(* IEC 61131-3 sources: iecf/harness/cases (part 4) *)

(* ---- bitarith.st ---- *)
(* Arithmetic on bit strings (the bit-string-arithmetic extension): a
   bit string counts as the unsigned integer of its width. Worked by
   hand, d 16#FFFF_FFF0, w 300, b 200, b2 100, i -5, x 513.7:
   %QD0  d + 16#20: DWORD, 16#1_0000_0010 wraps to 16#10, flagged.
   %QW4  w * 2 + b: WORD, 800 (16#0320); b widens to WORD.
   %QB6  b + b2: BYTE, 300 wraps to 44 (16#2C), flagged.
   %QW8  i + b: INT, -5 + 200 = 195; b counts as USINT, which INT holds.
   %QD12 BYTE_TO_REAL(b) + WORD_TO_REAL(w) / 3.0: 200.0 + 100.0 = 300.0
         (16#43960000), by value.
   %QB16 REAL_TO_BYTE(x / 10.0): 51.37 rounds to 51 (16#33).
   %QW18 w MOD 7 + b / 3: WORD 6 and BYTE 66 (division toward 0), as
         WORD 72 (16#48), into a UINT.
   %QB20 b - b2 * 2: 200 - 200 = 0.
   %QW22 a[b]: the array indexed by a BYTE, a[200] = 7.
   %QD24 DWORD_TO_REAL(16#3F800000) > 0.5: Ed.3's binary transfer is
         kept, 1.0 > 0.5, TRUE, 1.
   reference-skip: arithmetic on bit strings is CODESYS's, not IEC 61131-3. *)
PROGRAM main
  VAR
    d : DWORD := 16#FFFF_FFF0; w : WORD := 300; b : BYTE := 200; b2 : BYTE := 100;
    i : INT := -5; x : REAL := 513.7;
    a : ARRAY[0..255] OF INT;
  END_VAR
  VAR
    q0 AT %QD0 : DWORD; q1 AT %QW4 : WORD; q2 AT %QB6 : BYTE; q3 AT %QW8 : INT;
    q4 AT %QD12 : REAL; q5 AT %QB16 : BYTE; q6 AT %QW18 : UINT; q7 AT %QB20 : BYTE;
    q8 AT %QW22 : INT; q9 AT %QD24 : DWORD;
  END_VAR
  a[b] := 7;
  q0 := d + 16#20;
  q1 := w * 2 + b;
  q2 := b + b2;
  q3 := i + b;
  q4 := BYTE_TO_REAL(b) + WORD_TO_REAL(w) / 3.0;
  q5 := REAL_TO_BYTE(x / 10.0);
  q6 := w MOD 7 + b / 3;
  q7 := b - b2 * 2;
  q8 := a[b];
  q9 := DWORD_TO_REAL(16#3F800000) > 0.5;
END_PROGRAM

CONFIGURATION cf
  RESOURCE r ON x
    TASK tk(INTERVAL := T#10ms, PRIORITY := 1);
    PROGRAM p WITH tk : main;
  END_RESOURCE
END_CONFIGURATION

(* ---- bits.st ---- *)
(* Bit strings and BOOL: AND OR XOR NOT, the shifts and rotations, and
   BOOL expressions with short and full evaluation alike. *)
PROGRAM main
VAR
  x AT %IW0 : WORD;
  n AT %IB2 : BYTE;
  b0 AT %IX3.0 : BOOL;
  b1 AT %IX3.1 : BOOL;
  r_and AT %MW0 : WORD;
  r_or AT %MW2 : WORD;
  r_xor AT %MW4 : WORD;
  r_not AT %MW6 : WORD;
  r_shl AT %MW8 : WORD;
  r_shr AT %MW10 : WORD;
  r_rol AT %MW12 : WORD;
  r_ror AT %MW14 : WORD;
  r_dw AT %MD16 : DWORD;
  r_lw AT %ML20 : LWORD;
  r_by AT %MB28 : BYTE;
  q0 AT %QX0.0 : BOOL;
  q1 AT %QX0.1 : BOOL;
  q2 AT %QX0.2 : BOOL;
  q3 AT %QX0.3 : BOOL;
  q4 AT %QX0.4 : BOOL;
END_VAR
r_and := x AND 16#0FF0;
r_or := x OR 16#8001;
r_xor := x XOR 16#FFFF;
r_not := NOT x;
r_shl := SHL(x, BYTE_TO_INT(n));
r_shr := SHR(x, BYTE_TO_INT(n));
r_rol := ROL(x, BYTE_TO_INT(n));
r_ror := ROR(x, BYTE_TO_INT(n));
r_dw := ROL(WORD_TO_DWORD(x), 20);
r_lw := SHL(WORD_TO_LWORD(x), 48) OR 16#FF;
r_by := NOT n XOR 16#0F;
q0 := b0 AND b1;
q1 := b0 OR b1;
q2 := b0 XOR b1;
q3 := NOT b0 & b1;
q4 := (b0 OR NOT b1) AND x <> 0;
END_PROGRAM

CONFIGURATION plant
  RESOURCE r ON PLC
    TASK fast(INTERVAL := T#10ms, PRIORITY := 0);
    PROGRAM p WITH fast : main;
  END_RESOURCE
END_CONFIGURATION

(* ---- caseany.st ---- *)
(* CASE on a selector of any elementary type (Ed.3 7.3.3.3.3: "a
   variable of elementary data type", its labels "literals, enumerated
   values, or subranges" it can be compared with): BOOL, the bit
   strings, CHAR and WCHAR, STRING and WSTRING, REAL, TIME, DATE and
   TOD; labels that are literals, constants and subranges; a selector
   that is a FUNCTION with effects, called once. q[i] is the arm taken,
   9 for ELSE. Worked by hand:

   tick 0, n 1: b TRUE 1; w 16#2 1; bb 1 1; lw 1 ELSE 9; 'a' 1; "a" 1;
   'ab' 1; "ab" 1; 1.0 1; T#1s 1; the date 1; noon 1. calls 1 (Q12).
   tick 1, n 2: b FALSE 2; w 16#4, in 4..8, 2; bb 2 ELSE 9; lw 2 1; 'c'
   in 'b'..'d' 2; "z" in "y".."z" 2; 'cd', the constant, 2; "zz" 2; 2.5
   in 2.0..3.0 2; T#3s in the constant 2s..5s 2; June in February to
   December 2; 13:30 2. calls 2.
   tick 2, n 3: b TRUE 1; w 16#8 2; bb 3 1; lw 3 9; 'x' 9; "q" 9; 'zz'
   in 'x'..'zzzz' 3; "q" 9; -1.0 9; T#9s 9; 2021 9; 01:00 9. calls 3.
   reference-skip: CASE on anything but an integer or an enumeration:
   refused. *)
FUNCTION bump : STRING[4]
  VAR_INPUT s : STRING[4]; END_VAR
  VAR_EXTERNAL calls : USINT; END_VAR
  calls := calls + 1;
  bump := s;
END_FUNCTION
PROGRAM main
  VAR CONSTANT kc : CHAR := 'b'; ks : STRING[4] := 'cd'; kt : TIME := T#2s; END_VAR
  VAR_EXTERNAL calls : USINT; END_VAR
  VAR b : BOOL; w : WORD; bb : BYTE; c : CHAR; s : STRING[4]; r : REAL; t : TIME; d : DATE; wc : WCHAR; lw : LWORD; ws : WSTRING[4]; tod1 : TOD; n : USINT; END_VAR
  VAR q AT %QB0 : ARRAY [0..11] OF USINT; qc AT %QB12 : USINT; END_VAR
  n := n + 1;
  b := (n MOD 2) = 1;
  w := SHL(WORD#1, n);
  bb := USINT_TO_BYTE(n);
  lw := USINT_TO_LWORD(n);
  CASE n OF 1: c := 'a'; s := 'ab'; wc := "a"; ws := "ab"; r := 1.0; t := T#1s; d := D#2020-01-01; tod1 := TOD#12:00:00;
            2: c := 'c'; s := 'cd'; wc := "z"; ws := "zz"; r := 2.5; t := T#3s; d := D#2020-06-15; tod1 := TOD#13:30:00;
  ELSE c := 'x'; s := 'zz'; wc := "q"; ws := "q"; r := -1.0; t := T#9s; d := D#2021-01-01; tod1 := TOD#01:00:00;
  END_CASE;
  CASE b OF TRUE: q[0] := 1; FALSE: q[0] := 2; END_CASE;
  CASE w OF 16#0002: q[1] := 1; 16#0004..16#0008: q[1] := 2; ELSE q[1] := 3; END_CASE;
  CASE bb OF 16#01, 16#03: q[2] := 1; ELSE q[2] := 9; END_CASE;
  CASE lw OF 16#2: q[3] := 1; ELSE q[3] := 9; END_CASE;
  CASE c OF 'a': q[4] := 1; kc..'d': q[4] := 2; ELSE q[4] := 9; END_CASE;
  CASE wc OF "a": q[5] := 1; "y".."z": q[5] := 2; ELSE q[5] := 9; END_CASE;
  CASE bump(s) OF 'ab': q[6] := 1; ks: q[6] := 2; 'x'..'zzzz': q[6] := 3; ELSE q[6] := 9; END_CASE;
  CASE ws OF "ab": q[7] := 1; "zz": q[7] := 2; ELSE q[7] := 9; END_CASE;
  CASE r OF 1.0: q[8] := 1; 2.0..3.0: q[8] := 2; ELSE q[8] := 9; END_CASE;
  CASE t OF T#1s: q[9] := 1; kt..T#5s: q[9] := 2; ELSE q[9] := 9; END_CASE;
  CASE d OF D#2020-01-01: q[10] := 1; D#2020-02-01..D#2020-12-31: q[10] := 2; ELSE q[10] := 9; END_CASE;
  CASE tod1 OF TOD#12:00:00: q[11] := 1; TOD#13:00:00..TOD#14:00:00: q[11] := 2; ELSE q[11] := 9; END_CASE;
  qc := calls;
END_PROGRAM
CONFIGURATION c VAR_GLOBAL calls : USINT; END_VAR RESOURCE r ON PLC TASK t(INTERVAL := T#10ms, PRIORITY := 1); PROGRAM p WITH t : main; END_RESOURCE END_CONFIGURATION

(* ---- caselimits.st ---- *)
(* CASE subrange labels with a bound at the selector type's own limit:
   `0..5` on a USINT, `-128..-1` and `1..127` on a SINT, `0..255` on a
   USINT, all of it. Such a bound tests nothing, and its comparison is
   one C calls always true (-Wtype-limits): the generated C must still
   be strict-clean. Worked by hand, n and b counting 0, 1, 2 from tick 0,
   s -128, then -1, then 126:

   tick 0: n 0 in 0..5: Q0 01; s -128: Q1 01; b 0: Q2 01.
   tick 1: n 1: 01; s -1: 01; b 1: 01.
   tick 2: n 2: 01; s 126: Q1 03; 01. *)
PROGRAM main
  VAR n : USINT; s : SINT := -128; b : USINT; k : INT; END_VAR
  VAR q0 AT %QB0 : USINT; q1 AT %QB1 : USINT; q2 AT %QB2 : USINT; END_VAR
  CASE n OF 0..5: q0 := 1; ELSE q0 := 2; END_CASE;
  CASE s OF -128..-1: q1 := 1; 0: q1 := 2; 1..127: q1 := 3; END_CASE;
  CASE b OF 0..255: q2 := 1; END_CASE;
  n := n + 1;
  b := b + 1;
  k := k + 1;
  IF k = 1 THEN s := -1; ELSE s := 126; END_IF;
END_PROGRAM
CONFIGURATION c RESOURCE r ON PLC TASK t(INTERVAL := T#10ms, PRIORITY := 1); PROGRAM p WITH t : main; END_RESOURCE END_CONFIGURATION

(* ---- casenamed.st ---- *)
(* A named value as a CASE label (Ed.3 6.4.4.3, 7.3.3.3.3): a constant,
   its number compared with the selector's. Found in TcOpen, where it
   was E0032. Worked by hand:
   %QW0: d is eDist#Y (20): the label eDist#Y, 2.
   %QW2: n is eNum#Q (5): the label eNum#Q, 4.
   %QW4: d's number through its base type, 20.
   reference-skip: matiec has no named values with values given. *)
TYPE eDist : (X := 10, Y := 20, Z := 30); END_TYPE
TYPE eNum : INT (P := 1, Q := 5); END_TYPE

PROGRAM main
  VAR d : eDist := eDist#Y; n : eNum := eNum#Q; END_VAR
  VAR q0 AT %QW0 : INT; q1 AT %QW2 : INT; q2 AT %QW4 : INT; END_VAR
  CASE d OF
    eDist#X: q0 := 1;
    eDist#Y: q0 := 2;
  ELSE
    q0 := 3;
  END_CASE;
  CASE n OF
    eNum#P: q1 := 3;
    eNum#Q: q1 := 4;
  END_CASE;
  q2 := TO_INT(d);
END_PROGRAM

CONFIGURATION cf
  RESOURCE r ON x
    TASK tk(INTERVAL := T#10ms, PRIORITY := 1);
    PROGRAM p WITH tk : main;
  END_RESOURCE
END_CONFIGURATION

(* ---- codesysanyto.st ---- *)
(* CODESYS's and TwinCAT's ANY_TO_<type> (any-to): Ed.3's overloaded
   TO_<type>, as TcOpen's TcoRealToBytes and StringBuilder call it.
   Worked by hand, d + 1 and b + 1 each tick, d from 41, b from 7:
   %QW0 ANY_TO_INT(r * 2.0), r = ANY_TO_REAL(d): tick 0 d 42: 84;
   %QW2 ANY_TO_INT(ANY_TO_STRING(b) + '0' joined): b 7: '70': 70;
   %QW4 ANY_TO_INT(ANY_TO_BOOL(b - 7)): b 7: FALSE: 0.
   tick 1: d 43: 86; b 8: 80; 1.
   reference-skip: not IEC 61131-3. *)
PROGRAM main
  VAR d : DINT := 41; r : REAL; b : BYTE := 7; END_VAR
  VAR q0 AT %QW0 : INT; END_VAR
  VAR q1 AT %QW2 : INT; END_VAR
  VAR q2 AT %QW4 : INT; END_VAR
  d := d + 1;
  r := ANY_TO_REAL(d);
  q0 := ANY_TO_INT(r * 2.0);
  q1 := ANY_TO_INT(CONCAT(ANY_TO_STRING(b), '0'));
  q2 := ANY_TO_INT(ANY_TO_BOOL(b - 7));
  b := b + 1;
END_PROGRAM

CONFIGURATION cf
  RESOURCE r ON x
    TASK tk(INTERVAL := T#10ms, PRIORITY := 1);
    PROGRAM p WITH tk : main;
  END_RESOURCE
END_CONFIGURATION

(* ---- codesyschain.st ---- *)
(* Found in OSCAT BUILDING (BOILER): chained assignment, read right to
   left, each inner target read back (chained-assignment). Worked by hand:
   %QD0: r := x := 7 / 2: x is INT, 7 / 2 is 3, r gets 3.0, 16#40400000.
   %QW4: x, 3.
   %QW6, %QW8: q := arr[i] := y := 9, i 2: arr[2] 9, q 9.
   %QW10: inside IF, a := b := c := 5 then a + b + c: 15.
   reference-skip: not IEC 61131-3. *)
PROGRAM main
  VAR
    x : INT; y : SINT; i : INT := 2; arr : ARRAY[0..3] OF INT;
    a : INT; b : INT; c : INT;
  END_VAR
  VAR
    r AT %QD0 : REAL; qx AT %QW4 : INT; q AT %QW6 : INT; q2 AT %QW8 : INT;
    q3 AT %QW10 : INT;
  END_VAR
  r := x := 7 / 2;
  qx := x;
  q := arr[i] := y := 9;
  q2 := arr[2];
  IF i = 2 THEN
    a := b := c := 5;
  END_IF;
  q3 := a + b + c;
END_PROGRAM

CONFIGURATION cf
  RESOURCE r ON x
    TASK tk(INTERVAL := T#10ms, PRIORITY := 1);
    PROGRAM p WITH tk : main;
  END_RESOURCE
END_CONFIGURATION

(* ---- codesysdates.st ---- *)
(* Found in OSCAT NETWORK and BUILDING, each an extension. Worked by hand:
   %QB0 bit 0: UDINT 70000 > DWORD 16#10000 (65536): a bit string compared
   with an integer, as its unsigned integer (bit-string-arithmetic): TRUE.
   %QB0 bit 1: BYTE 200 < INT 100: FALSE.
   %QW2: TOD_TO_TIME(TOD#01:00:00) is T#1h, as DINT ms / 1000, 3600.
   %QD4: TIME_TO_TOD(T#1d2h3m4s5ms) drops the day: TOD#02:03:04.005,
   7384005 ms (date-number-conversions).
   %QD8: D#2026-11-19 + T#1d - T#2d is D#2026-11-18; DATE_TO_UDINT /
   86400 counts its days since 1970-01-01: 20775
   (date-time-arithmetic).
   %QB12: d2 := d + half, half T#12h a variable: no whole day, flagged
   and left undone, d2 stays D#1970-01-01: DATE_TO_UDINT(d2) = 0.
   reference-skip: none of these is IEC 61131-3. *)
PROGRAM main
  VAR
    u : UDINT := 70000; w : DWORD := 16#10000; b : BYTE := 200; i : INT := 100;
    d : DATE := D#2026-11-19; d2 : DATE; half : TIME := T#12h;
  END_VAR
  VAR
    x0 AT %QX0.0 : BOOL; x1 AT %QX0.1 : BOOL; q1 AT %QW2 : INT; q2 AT %QD4 : UDINT;
    q3 AT %QD8 : UDINT; q4 AT %QB12 : BYTE;
  END_VAR
  x0 := u > w;
  x1 := b < i;
  q1 := DINT_TO_INT(TIME_TO_DINT(TOD_TO_TIME(TOD#01:00:00)) / 1000);
  q2 := TOD_TO_UDINT(TIME_TO_TOD(T#1d2h3m4s5ms));
  q3 := DATE_TO_UDINT(d + T#1d - T#2d) / 86400;
  d2 := d + half;
  q4 := UDINT_TO_BYTE(DATE_TO_UDINT(d2));
END_PROGRAM

CONFIGURATION cf
  RESOURCE r ON x
    TASK tk(INTERVAL := T#10ms, PRIORITY := 1);
    PROGRAM p WITH tk : main;
  END_RESOURCE
END_CONFIGURATION

(* ---- codesysdtliterals.st ---- *)
(* A DT literal's seconds left out, and a fraction of its second
   (dt-literals): the seconds 0, the fraction dropped, W0016 - as
   TcOpen's TcoMessenger writes DT#1970-01-01-00:00 and its
   fbManipulatorAutomat DT#2013-05-09-13:29:20.500. Worked by hand,
   each as its seconds since 1970 (date-number-conversions):
   DT#1970-01-01-00:01: 60, 16#3C (%QD0).
   DT#2013-05-09-13:29:20.500: 2013-05-09 is day 15834, 1368057600 s;
   13:29:20 is 48560 s; 1368106160, 16#518BA4B0 (%QD4).
   An initial value DT#1970-01-02-00:00:00.999: one day, 86400, 16#15180
   (%QD8).
   reference-skip: not IEC 61131-3. *)
PROGRAM main
  VAR
    a : DT; b : DT; c : DT := DT#1970-01-02-00:00:00.999;
  END_VAR
  VAR q0 AT %QD0 : UDINT; q1 AT %QD4 : UDINT; q2 AT %QD8 : UDINT; END_VAR
  a := DT#1970-01-01-00:01;
  b := DT#2013-05-09-13:29:20.500;
  q0 := DT_TO_UDINT(a);
  q1 := DT_TO_UDINT(b);
  q2 := DT_TO_UDINT(c);
END_PROGRAM

CONFIGURATION cf
  RESOURCE r ON x
    TASK tk(INTERVAL := T#10ms, PRIORITY := 1);
    PROGRAM p WITH tk : main;
  END_RESOURCE
END_CONFIGURATION

(* ---- codesysenum.st ---- *)
(* CODESYS's enumerations (the codesys-enums extension,
   docs/extensions.md): the base type after the values, `(...) DWORD :=
   black`, and a value named `COLOR.green`, as CODESYS and TwinCAT write
   them (their `qualified_only` makes every use so); the attributes
   before a TYPE are pragmas, which iecf reads past. Worked by hand:
   COLOR is DWORD, black its initial value: c is 16#88000000, its top
   byte 16#88 (%QB0); c := COLOR.green, 16#FF00FF00, top byte 16#FF
   (%QB1); c = COLOR.green TRUE (%QX4.0). Lib.Mode (stop, run, fault)
   starts as Lib.Mode.stop: m = Lib.Mode.stop, 1 at tick 0, then 0
   (%QB2); m := Lib.Mode.run; CASE m OF Lib.Mode.run: %QB3 := 7.
   reference-skip: CODESYS's writing is not IEC 61131-3. *)
{attribute 'qualified_only'}
{attribute 'strict'}
TYPE COLOR :
(
    white := 16#FFFFFF00,
    green := 16#FF00FF00,
    black := 16#88000000
) DWORD := black
;
END_TYPE

NAMESPACE Lib
  TYPE Mode : (stop, run, fault); END_TYPE
END_NAMESPACE

PROGRAM main
  VAR c : COLOR; m : Lib.Mode := Lib.Mode.stop; END_VAR
  VAR
    q0 AT %QB0 : BYTE;
    q1 AT %QB1 : BYTE;
    q2 AT %QB2 : SINT;
    q3 AT %QB3 : SINT;
    b0 AT %QX4.0 : BOOL;
  END_VAR
  c := COLOR#black;
  q0 := DWORD_TO_BYTE(SHR(c, 24));
  c := COLOR.green;
  q1 := DWORD_TO_BYTE(SHR(c, 24));
  b0 := c = COLOR.green;
  q2 := SEL(m = Lib.Mode.stop, SINT#0, SINT#1);
  m := Lib.Mode.run;
  CASE m OF
    Lib.Mode.stop: q3 := 1;
    Lib.Mode.run: q3 := 7;
  END_CASE;
END_PROGRAM

CONFIGURATION cf
  RESOURCE r ON x
    TASK t(INTERVAL := T#10ms, PRIORITY := 1);
    PROGRAM p WITH t : main;
  END_RESOURCE
END_CONFIGURATION

(* ---- codesysgvl.st ---- *)
(* Global variable lists (--gvl, --qualified-gvl), as CODESYS and TwinCAT
   name them: IO (codesysgvl.d/io.st) and CFG, qualified-only
   (codesysgvl.d/cfg.st). Worked by hand:
   cycle 0: %QW0 IO.a + CFG.k = 3 + 7 = 10; r[CFG.N] := IO.a, %QW2 3;
     IO.a 4, read bare: %QW4 4; CFG.t[4] := 4 + 1, %QW6 5.
   cycle 1: 4 + 7 = 11; 4; 5; 6.
   reference-skip: not IEC 61131-3. *)
PROGRAM main
  VAR r : ARRAY[1..CFG.N] OF INT; END_VAR
  VAR x AT %QW0 : INT; y AT %QW2 : INT; z AT %QW4 : INT; w AT %QW6 : INT; END_VAR
  x := IO.a + CFG.k;
  r[CFG.N] := IO.a;
  y := r[4];
  IO.a := IO.a + 1;
  z := a;
  CFG.t[CFG.N] := a + 1;
  w := CFG.t[4];
END_PROGRAM

CONFIGURATION cf
  RESOURCE r ON x
    TASK tk(INTERVAL := T#10ms, PRIORITY := 1);
    PROGRAM p WITH tk : main;
  END_RESOURCE
END_CONFIGURATION

(* ---- codesysjump.st ---- *)
(* Found in OSCAT NETWORK (IP_CONTROL2): JMP and labels in ST
   (jump-labels). Worked by hand:
   %QW0: i counted to 5 by a jump back: 5.
   %QW2: JMP out of the FOR at k = 3, k left as the body has it: 3.
   %QW4: n = 1 + 2 + 3: 6; the jumped-over q2 := 99 never runs.
   %QW6: arr[k] with k 2 holds; k 7 on the jump back is outside 0..3:
   INDEX fault on the line of arr[k] := 1 (32), the task stops: q3 1.
   reference-skip: not IEC 61131-3. *)
PROGRAM main
  VAR i : INT; k : INT; n : INT; arr : ARRAY[0..3] OF INT; END_VAR
  VAR q0 AT %QW0 : INT; q1 AT %QW2 : INT; q2 AT %QW4 : INT; q3 AT %QW6 : INT; END_VAR
  i := 0;
  n := 0;
again:
  i := i + 1;
  IF i < 5 THEN
    JMP again;
  END_IF;
  q0 := i;
  JMP skip;
  q2 := 99;
skip:
  FOR k := 1 TO 10 DO
    n := n + k;
    IF k = 3 THEN JMP out; END_IF;
  END_FOR;
out:
  q1 := k;
  q2 := n;
  k := 2;
back:
  arr[k] := 1;
  k := k + 5;
  q3 := q3 + 1;
  IF k < 20 THEN JMP back; END_IF;
END_PROGRAM

CONFIGURATION cf
  RESOURCE r ON x
    TASK tk(INTERVAL := T#10ms, PRIORITY := 1);
    PROGRAM p WITH tk : main;
  END_RESOURCE
END_CONFIGURATION

(* ---- codesyslibprograms.st ---- *)
(* A library's PROGRAMs in its namespace, as CODESYS and TwinCAT have
   them: the library A (codesyslibprograms.d/a.st) and B, qualified-only
   (b.st), each with a MAIN of its own, beside this project's MAIN. A's
   Counter is called and read by its short name, through A's USING,
   from here and from A's own block User, and its method called;
   A.MAIN and B.MAIN by the library's name (program-instances).
   Worked by hand:
   cycle 0: Counter() v 10, %QW0 10; A.MAIN() n 1, %QW2 1; B.MAIN()
     x 100, %QW4 100; u(), Counter() again, %QW6 20; A.Counter.Bump(5),
     %QW8 25.
   cycle 1: 35; 2; 200; 45; 50.
   reference-skip: not IEC 61131-3. *)
PROGRAM MAIN
  VAR u : User; END_VAR
  VAR q0 AT %QW0 : INT; q1 AT %QW2 : INT; q2 AT %QW4 : INT; q3 AT %QW6 : INT; q4 AT %QW8 : INT; END_VAR
  Counter();
  q0 := Counter.v;
  A.MAIN();
  q1 := A.MAIN.n;
  B.MAIN();
  q2 := B.MAIN.x;
  u();
  q3 := Counter.v;
  A.Counter.Bump(5);
  q4 := A.Counter.v;
END_PROGRAM

CONFIGURATION cf
  RESOURCE r ON x
    TASK tk(INTERVAL := T#10ms, PRIORITY := 1);
    PROGRAM p WITH tk : MAIN;
  END_RESOURCE
END_CONFIGURATION

(* ---- codesysliteralwidening.st ---- *)
(* An untyped integer literal the other operand's type does not hold
   (literal-widening): the operation is computed in the narrowest type
   of the operand's kind that holds it, as CODESYS and TwinCAT compute
   intermediate results at least 32 bits wide. TcOpen's TcoBytesToReal
   writes `256 * _b0 + _b1` of BYTEs and `w * 65536` of a WORD, its
   TcoRealToBytes `2147483648 + ...` of DINTs.
   Worked by hand:
   256 * 16#12 + 16#34, in WORD: 16#1234 (4660).
   16#0003 * 65536 + 16#1234, in DWORD: 16#00031234 (201268).
   2147483648 + 100, in LINT: 2147483748 (16#80000064).
   5 * -1 of a UINT, in DINT: -5.
   30000 < 70000 of an INT, compared in DINT: TRUE.
   reference-skip: not IEC 61131-3. *)
PROGRAM main
  VAR
    b0 : BYTE := 16#12;
    b1 : BYTE := 16#34;
    w : WORD;
    w1 : WORD := 16#0003;
    k : INT := 30000;
    x : DINT := 100;
    u : UINT := 5;
  END_VAR
  VAR q0 AT %QD0 : DWORD; q4 AT %QD4 : DWORD; q8 AT %QL8 : LINT; q16 AT %QD16 : DINT; q20 AT %QX20.0 : BOOL; END_VAR
  w := 256 * b0 + b1;
  q0 := w;
  q4 := (w1 * 65536) + w;
  q8 := 2147483648 + x;
  q16 := u * -1;
  q20 := k < 70000;
END_PROGRAM

CONFIGURATION cf
  RESOURCE r ON x
    TASK tk(INTERVAL := T#10ms, PRIORITY := 1);
    PROGRAM p WITH tk : main;
  END_RESOURCE
END_CONFIGURATION

(* ---- codesyspack.st ---- *)
(* The codesys pack (docs/extensions.md, "Packs"): one name for the
   extensions code written for CODESYS and TwinCAT uses, seven of them
   here. Worked by hand:
   gCount, a top-level global, used without VAR_EXTERNAL
   (implicit-externals) and bound to a REFERENCE TO (reference-to): r :=
   r + 1 makes it 6, then 7 (%QB3). t T#1500ms; ms := TIME_TO_DINT(t),
   1500 (time-number-conversions), worked out as it is set up
   (initial-expressions): ms / 100, 15 (%QB0). Len3 takes a VAR_IN_OUT
   CONSTANT STRING(10) (in-out-constant, string-parentheses), given 16
   characters, all of them read: n := Len3('abcdefghijklmnop') + ms,
   1516; n - 1500, 16 (%QB1). m : E_Mode := E_Mode.eRun, its base type
   after its values (codesys-enums): m = E_Mode.eRun, 1 (%QB2).
   BYTE_TO_BOOL(16#10) TRUE (bit-string-to-bool, %QX4.0).
   reference-skip: CODESYS's extensions are not IEC 61131-3. *)
VAR_GLOBAL gCount : INT := 5; END_VAR

TYPE E_Mode : (eIdle, eRun) DWORD; END_TYPE

FUNCTION Len3 : DINT
  VAR_IN_OUT CONSTANT s : STRING(10); END_VAR
  Len3 := INT_TO_DINT(LEN(s));
END_FUNCTION

PROGRAM main
  VAR
    t : TIME := T#1500ms;
    ms : DINT := TIME_TO_DINT(t);
    n : DINT := Len3('abcdefghijklmnop') + ms;
    m : E_Mode := E_Mode.eRun;
    r : REFERENCE TO INT;
    b : BOOL := BYTE_TO_BOOL(16#10);
  END_VAR
  VAR
    q0 AT %QB0 : SINT;
    q1 AT %QB1 : SINT;
    q2 AT %QB2 : SINT;
    q3 AT %QB3 : SINT;
    b0 AT %QX4.0 : BOOL;
  END_VAR
  r REF= gCount;
  r := r + 1;
  q0 := DINT_TO_SINT(ms / 100);
  q1 := DINT_TO_SINT(n - 1500);
  q2 := SEL(m = E_Mode.eRun, SINT#0, SINT#1);
  q3 := INT_TO_SINT(gCount);
  b0 := b;
END_PROGRAM

CONFIGURATION cf
  RESOURCE r ON x
    TASK tk(INTERVAL := T#10ms, PRIORITY := 1);
    PROGRAM p WITH tk : main;
  END_RESOURCE
END_CONFIGURATION

(* ---- codesyssemi.st ---- *)
(* Found in TcOpen (TwinCAT), 10639 ends without ';' against 829 with,
   and in OSCAT: END_IF and its kin with no ';' (optional-semicolons).
   Worked by hand:
   %QW0: n counts 1 + 2 + 3 + 4 by FOR, then +10 by IF: 20.
   %QW2: WHILE doubles w from 1 past 100: 128; REPEAT halves it to 64,
   then CASE adds 1 for 64: 65.
   reference-skip: not IEC 61131-3. *)
PROGRAM main
  VAR n : INT; i : INT; w : INT := 1; END_VAR
  VAR q0 AT %QW0 : INT; q1 AT %QW2 : INT; END_VAR
  n := 0;
  FOR i := 1 TO 4 DO
    n := n + i;
  END_FOR
  IF n = 10 THEN
    n := n + 10;
  END_IF
  WHILE w <= 100 DO
    w := w * 2;
  END_WHILE
  REPEAT
    w := w / 2;
  UNTIL w <= 100 END_REPEAT
  CASE w OF
    64: w := w + 1;
  END_CASE
  q0 := n;
  q1 := w;
END_PROGRAM

CONFIGURATION cf
  RESOURCE r ON x
    TASK tk(INTERVAL := T#10ms, PRIORITY := 1);
    PROGRAM p WITH tk : main;
  END_RESOURCE
END_CONFIGURATION

(* ---- codesysstraysemi.st ---- *)
(* A `;` that ends nothing (stray-semicolons), as TcOpen writes
   `END_TYPE;` after its EtherCAT structures and `p : T;;` in a VAR
   section; END_PROGRAM; too: dropped, the declarations read as
   without it.
   Worked by hand, each tick: s.a + 1 and s.b + 2 from 0; k counts.
   Tick 1: 1, 2, 1; tick 2: 2, 4, 2.
   reference-skip: not IEC 61131-3. *)
TYPE Pair :
STRUCT
  a : INT;
  b : INT;
END_STRUCT
END_TYPE;

PROGRAM main
  VAR
    s : Pair;;
    ;
    k : INT;
  END_VAR
  VAR q0 AT %QW0 : INT; q2 AT %QW2 : INT; q4 AT %QW4 : INT; END_VAR
  s.a := s.a + 1;
  s.b := s.b + 2;
  k := k + 1;
  q0 := s.a;
  q2 := s.b;
  q4 := k;
END_PROGRAM;

CONFIGURATION cf
  RESOURCE r ON x
    TASK tk(INTERVAL := T#10ms, PRIORITY := 1);
    PROGRAM p WITH tk : main;
  END_RESOURCE
END_CONFIGURATION

(* ---- codesysstructext.st ---- *)
(* A structure extending another (struct-extends), as TcOpen's I/O types
   do: TYPE X EXTENDS Base : STRUCT, the base's fields first, at any
   depth, their initial values with them. Worked by hand:
   %QW0: t.a := 1, then a + b + c + d: 1 + 2 + 3 + 4 = 10.
   %QW2: a Top given to a Middle's field by field: Middle.c, 3.
   reference-skip: not IEC 61131-3. *)
TYPE
  Base : STRUCT a : INT; b : INT := 2; END_STRUCT;
  Middle EXTENDS Base : STRUCT c : INT := 3; END_STRUCT;
  Top EXTENDS Middle : STRUCT d : INT := 4; END_STRUCT;
END_TYPE

PROGRAM main
  VAR t : Top; m : Middle; END_VAR
  VAR q AT %QW0 : INT; r AT %QW2 : INT; END_VAR
  t.a := 1;
  q := t.a + t.b + t.c + t.d;
  m.c := t.c;
  r := m.c;
END_PROGRAM

CONFIGURATION cf
  RESOURCE r ON x
    TASK tk(INTERVAL := T#10ms, PRIORITY := 1);
    PROGRAM p WITH tk : main;
  END_RESOURCE
END_CONFIGURATION

(* ---- codesyssyntax.st ---- *)
(* Three CODESYS ways of writing, each an extension (docs/extensions.md).
   Worked by hand:
   struct-semicolon: Pair ends END_STRUCT with no ';', the next type
   follows; Trio's END_STRUCT stands before END_TYPE.
   bare-array-init: a : ARRAY[1..5] OF SINT := 1, 2, 2(7), 3; is
   [1, 2, 7, 7, 3], sum 20 (%QB0); Pair's v := 8, 9 in a STRUCT, 8 + 9 =
   17 (%QB1); the type Row := 4, 5, 6, 4 + 5 + 6 = 15 (%QB2).
   real-without-point: r := 1E3 + 25E-1, 1002.5; REAL_TO_SINT(r / 100.0)
   is 10.025 rounded, 10 (%QB3); Trio's z := 2E1, 20.0, as SINT 20
   (%QB4).
   reference-skip: none of the three is IEC 61131-3. *)
TYPE
  Pair : STRUCT
    v : ARRAY[1..2] OF SINT := 8, 9;
  END_STRUCT
  Row : ARRAY[0..2] OF SINT := 4, 5, 6;
  Trio : STRUCT
    z : REAL := 2E1;
  END_STRUCT
END_TYPE

PROGRAM main
  VAR
    a : ARRAY[1..5] OF SINT := 1, 2, 2(7), 3;
    p : Pair;
    w : Row;
    t : Trio;
    r : REAL;
    i : INT;
    s : SINT;
  END_VAR
  VAR
    q0 AT %QB0 : SINT;
    q1 AT %QB1 : SINT;
    q2 AT %QB2 : SINT;
    q3 AT %QB3 : SINT;
    q4 AT %QB4 : SINT;
  END_VAR
  s := 0;
  FOR i := 1 TO 5 DO
    s := s + a[i];
  END_FOR;
  q0 := s;
  q1 := p.v[1] + p.v[2];
  q2 := w[0] + w[1] + w[2];
  r := 1E3 + 25E-1;
  q3 := REAL_TO_SINT(r / 100.0);
  q4 := REAL_TO_SINT(t.z);
END_PROGRAM

CONFIGURATION cf
  RESOURCE r ON x
    TASK tk(INTERVAL := T#10ms, PRIORITY := 1);
    PROGRAM p WITH tk : main;
  END_RESOURCE
END_CONFIGURATION

(* ---- codesysunion.st ---- *)
(* CODESYS's and TwinCAT's UNION (union), as a STRUCT OVERLAP whose every
   member is AT %B0: un set up through d alone, 1.0's bits (16#3F800000);
   r, declared first, is not defaulted over it. Worked by hand:
   %QD0: q := un.r before un.r is changed, 1.0's bytes, 00 00 80 3f.
   un.r := 2.0 changes the same bytes un.d reads.
   %QD4: w := un.d after that, 2.0's bits read as a DWORD, 00 00 00 40.
   reference-skip: not IEC 61131-3. *)
TYPE
  U : UNION
    r : REAL;
    d : DWORD;
  END_UNION;
END_TYPE

PROGRAM main
  VAR un : U := (d := 16#3F800000); END_VAR
  VAR q AT %QD0 : REAL; w AT %QD4 : DWORD; END_VAR
  q := un.r;
  un.r := 2.0;
  w := un.d;
END_PROGRAM

CONFIGURATION cf
  RESOURCE r ON x
    TASK tk(INTERVAL := T#10ms, PRIORITY := 1);
    PROGRAM p WITH tk : main;
  END_RESOURCE
END_CONFIGURATION

(* ---- connections.st ---- *)
(* Program connections (Ed.3 6.8.2): a program instance's inputs given a
   literal, a global or an address, its outputs written to a global or an
   address. Each input is set before the instance runs, each output
   taken after it. The reference compiler crashes on a literal input and writes C that
   does not compile for the rest (PROPOSAL.md §1b): the trace is iecf's
   alone, connections.iecf.trace, checked by hand.

   Instance a adds 1 a tick, b adds the global ten (10), c the input
   global k (at %IW0). a's total goes to the global sum, b's to the
   global out_b (at %MD4), c's to out_c (at %MD8); a's done, inverted,
   straight to the address %QX0.0, a bare BOOL. *)
PROGRAM counter
VAR_INPUT inc : INT; END_VAR
VAR_OUTPUT total : DINT; done : BOOL; END_VAR
total := total + inc;
done := total >= 3;
END_PROGRAM

PROGRAM report
VAR_EXTERNAL sum : DINT; END_VAR
VAR r_sum AT %MD0 : DINT; END_VAR
r_sum := sum;
END_PROGRAM

CONFIGURATION plant
  VAR_GLOBAL
    ten : INT := 10;
    sum : DINT;
  END_VAR
  VAR_GLOBAL
    k AT %IW0 : INT;
    out_b AT %MD4 : DINT;
    out_c AT %MD8 : DINT;
  END_VAR
  RESOURCE r ON PLC
    TASK fast(INTERVAL := T#10ms, PRIORITY := 0);
    PROGRAM a WITH fast : counter(inc := 1, total => sum, NOT done => %QX0.0);
    PROGRAM b WITH fast : counter(inc := ten, total => out_b);
    PROGRAM c WITH fast : counter(inc := k, total => out_c);
    PROGRAM rep WITH fast : report;
  END_RESOURCE
END_CONFIGURATION

(* ---- conrefs.st ---- *)
(* Program connections (Ed.3 6.8.2) of a reference, in and out, and of
   NULL; a CHAR output into a STRING global and a WCHAR one into a
   WSTRING global (Figure 11, implicit). The three programs run in
   order on one task. Worked by hand: setup points gr at gi (5). p1 gets
   gr, adds 1 to what it references and gives it back as ro, into gro;
   p2 gets NULL and does nothing, its ro NULL into gro2. Tick 0: gi 6
   (%QB0), gro^ 6 (%QB1), gro2 NULL (%QX2.0), gs 'k' (%QX2.1), gws "z"
   (%QX2.2). Tick 1: gi 7, gro^ 7.
   reference-skip: program connections, as connections; and REF_TO. *)
PROGRAM setup
  VAR_EXTERNAL gi : INT; gr : REF_TO INT; END_VAR
  gr := REF(gi);
END_PROGRAM

PROGRAM prod
  VAR_INPUT r : REF_TO INT; END_VAR
  VAR_OUTPUT ro : REF_TO INT; c : CHAR; wc : WCHAR; END_VAR
  IF r <> NULL THEN
    r^ := r^ + 1;
  END_IF;
  ro := r;
  c := 'k';
  wc := WCHAR#"z";
END_PROGRAM

PROGRAM show
  VAR_EXTERNAL gi : INT; gro, gro2 : REF_TO INT; gs : STRING[4]; gws : WSTRING[4]; END_VAR
  VAR
    q0 AT %QB0 : SINT;
    q1 AT %QB1 : SINT;
    b0 AT %QX2.0 : BOOL;
    b1 AT %QX2.1 : BOOL;
    b2 AT %QX2.2 : BOOL;
  END_VAR
  q0 := INT_TO_SINT(gi);
  IF gro <> NULL THEN
    q1 := INT_TO_SINT(gro^);
  END_IF;
  b0 := gro2 = NULL;
  b1 := gs = 'k';
  b2 := gws = "z";
END_PROGRAM

CONFIGURATION cf
  VAR_GLOBAL
    gi : INT := 5;
    gr, gro, gro2 : REF_TO INT;
    gs : STRING[4];
    gws : WSTRING[4];
  END_VAR
  RESOURCE r ON PLC
    TASK t(INTERVAL := T#10ms, PRIORITY := 1);
    PROGRAM s WITH t : setup;
    PROGRAM p1 WITH t : prod(r := gr, ro => gro, c => gs, wc => gws);
    PROGRAM p2 WITH t : prod(r := NULL, ro => gro2);
    PROGRAM v WITH t : show;
  END_RESOURCE
END_CONFIGURATION

(* ---- constinit2.st ---- *)
(* Initial values that are functions of constants (Table 34's string
   functions, the conversions of whole numbers to and from text, Tables
   30 and 36's date functions): worked out by the compiler. Each is
   compared with the same function of variables, computed as the program
   runs; ok counts those that agree, 19 of 19 (Q0 13). Worked by hand
   for three: LEN of s6, 'abZZef', is 6 (Q1); f1, FIND('abcabc', 'ca'),
   is 3 (Q2); i1, STRING_TO_INT('17'), is 17 (Q3 11).
   reference-skip: the reference compiler takes a literal there. *)
PROGRAM main
  VAR CONSTANT pre : STRING[4] := 'ab'; END_VAR
  VAR
    s1 : STRING[8] := CONCAT('ab', 'cd');
    s2 : STRING[8] := CONCAT(pre, '-x', 'y');
    l1 : INT := LEN('hello');
    s3 : STRING[8] := INT_TO_STRING(-42);
    s4 : STRING[8] := LEFT('abcdef', 3);
    s5 : STRING[8] := RIGHT('abcdef', 2);
    s6 : STRING[8] := REPLACE('abcdef', 'ZZ', 2, 3);
    s7 : STRING[8] := MID('abcdef', 2, 3);
    s9 : STRING[8] := INSERT('abcd', 'XY', 2);
    s10 : STRING[8] := DELETE('abcdef', 2, 3);
    ws : WSTRING[8] := CONCAT("ab", "cd");
    f1 : INT := FIND('abcabc', 'ca');
    i1 : INT := STRING_TO_INT('17');
    d1 : DATE := CONCAT_DATE(2020, 2, 29);
    dt1 : DT := CONCAT_DATE_TOD(D#2020-01-01, TOD#12:00:00);
    t3 : TIME := SUB_TOD_TOD(TOD#10:00:00, TOD#09:00:00);
    d3 : DT := ADD_DT_TIME(DT#2021-05-06-07:08:09, T#1h);
    tod1 : TOD := CONCAT_TOD(1, 2, 3, 4);
    dt2 : DT := CONCAT_DT(2020, 1, 1, 12, 0, 0, 0);
  END_VAR
  VAR a : STRING[8] := 'abcdef'; b : STRING[8] := 'ab'; c : STRING[8] := 'cd'; z : STRING[8] := 'ZZ'; n42 : INT := -42;
      two : INT := 2; three : INT := 3; y : INT := 2020; wa : WSTRING[8] := "ab"; wc : WSTRING[8] := "cd";
      dd : DATE := D#2020-01-01; tt : TOD := TOD#12:00:00; ta : TOD := TOD#10:00:00; tb : TOD := TOD#09:00:00;
      dx : DT := DT#2021-05-06-07:08:09; h : TIME := T#1h; ok : USINT; s17 : STRING[8] := '17'; abc2 : STRING[8] := 'abcabc';
      ca : STRING[8] := 'ca'; xy : STRING[8] := 'XY'; abcd : STRING[8] := 'abcd'; one : INT := 1; four : INT := 4; twelve : INT := 12; zero : INT;
  END_VAR
  VAR q AT %QB0 : USINT; q1 AT %QB1 : USINT; q2 AT %QB2 : USINT; q3 AT %QB3 : USINT; END_VAR
  ok := 0;
  IF s1 = CONCAT(b, c) THEN ok := ok + 1; END_IF;
  IF s2 = CONCAT(b, '-x', 'y') THEN ok := ok + 1; END_IF;
  IF l1 = LEN(CONCAT('hel', 'lo')) THEN ok := ok + 1; END_IF;
  IF s3 = INT_TO_STRING(n42) THEN ok := ok + 1; END_IF;
  IF s4 = LEFT(a, three) THEN ok := ok + 1; END_IF;
  IF s5 = RIGHT(a, two) THEN ok := ok + 1; END_IF;
  IF s6 = REPLACE(a, z, two, three) THEN ok := ok + 1; END_IF;
  IF s7 = MID(a, two, three) THEN ok := ok + 1; END_IF;
  IF s9 = INSERT(abcd, xy, two) THEN ok := ok + 1; END_IF;
  IF s10 = DELETE(a, two, three) THEN ok := ok + 1; END_IF;
  IF ws = CONCAT(wa, wc) THEN ok := ok + 1; END_IF;
  IF f1 = FIND(abc2, ca) THEN ok := ok + 1; END_IF;
  IF i1 = STRING_TO_INT(s17) THEN ok := ok + 1; END_IF;
  IF d1 = CONCAT_DATE(y, two, 29) THEN ok := ok + 1; END_IF;
  IF dt1 = CONCAT_DATE_TOD(dd, tt) THEN ok := ok + 1; END_IF;
  IF t3 = SUB_TOD_TOD(ta, tb) THEN ok := ok + 1; END_IF;
  IF d3 = ADD_DT_TIME(dx, h) THEN ok := ok + 1; END_IF;
  IF tod1 = CONCAT_TOD(one, two, three, four) THEN ok := ok + 1; END_IF;
  IF dt2 = CONCAT_DT(y, one, one, twelve, zero, zero, zero) THEN ok := ok + 1; END_IF;
  q := ok;
  q1 := INT_TO_USINT(LEN(s6));
  q2 := INT_TO_USINT(f1);
  q3 := INT_TO_USINT(i1);
END_PROGRAM
CONFIGURATION c RESOURCE r ON PLC TASK t(INTERVAL := T#10ms, PRIORITY := 1); PROGRAM p WITH t : main; END_RESOURCE END_CONFIGURATION

(* ---- constinit3.st ---- *)
(* More initial values worked out by the compiler, each compared with
   the same expression of variables computed as the program runs: + and
   - on dates (Table 35, a TOD wrapping at midnight), the long dates'
   functions, the text of a real, a duration and a date (the target's,
   written at start-up), a literal's text to its value, and reals that
   go through the target's mathematics to an integer away from where the
   conversion changes (docs/dependencies.md). ok counts those that
   agree, 24 of 24 (Q0 18). Worked by hand for three: x1, REAL_TO_INT
   of SQRT(16.0), is 4 (Q1); x5, 100 / x1, 25 (Q2 19); t3, TOD#23:00:00
   + T#2h, is 01:00, its hour 1 (Q3).
   reference-skip: the reference compiler takes a literal there. *)
PROGRAM main
  VAR
    d5 : DT := DT#2021-05-06-07:08:09 + T#1h;
    d6 : DT := DT#2021-05-06-07:08:09 - T#1h;
    t1 : TIME := DT#2021-05-06-07:08:09 - DT#2021-05-06-07:00:00;
    t2 : TIME := D#2021-05-07 - D#2021-05-06;
    t3 : TOD := TOD#23:00:00 + T#2h;
    t4 : TIME := TOD#10:00:00 - TOD#09:00:00;
    l1 : LDT := LDT#2021-05-06-07:08:09 + LT#1h;
    l2 : LTIME := LDT#2021-05-06-07:08:09 - LDT#2021-05-06-07:00:00;
    l3 : LTOD := CONCAT_LTOD(1, 2, 3, 4);
    l4 : LDT := CONCAT_LDT(2020, 1, 1, 12, 0, 0, 0);
    l5 : LDT := CONCAT_DATE_LTOD(D#2020-01-01, LTOD#12:00:00);
    l6 : LTOD := ADD_LTOD_LTIME(LTOD#23:00:00, LT#2h);
    s1 : STRING[30] := REAL_TO_STRING(1.5);
    s3 : STRING[40] := TIME_TO_STRING(T#1h30m);
    s4 : STRING[24] := DT_TO_STRING(DT#2021-05-06-07:08:09);
    r1 : REAL := STRING_TO_REAL('1.5');
    tm : TIME := STRING_TO_TIME('T#5s');
    dd : DATE := STRING_TO_DATE('D#2021-05-06');
    b1 : BOOL := STRING_TO_BOOL('TRUE');
    x1 : INT := REAL_TO_INT(SQRT(16.0));
    x3 : INT := REAL_TO_INT(SQRT(2.0) * 100.0);
    x4 : REAL := 10.0 / SQRT(2.0);
    x5 : INT := 100 / REAL_TO_INT(SQRT(16.0));
    x11 : DINT := LREAL_TO_DINT(1.0E5 * SQRT(LREAL#2.0));
  END_VAR
  VAR dx : DT := DT#2021-05-06-07:08:09; dy : DT := DT#2021-05-06-07:00:00; h : TIME := T#1h; h2 : TIME := T#2h;
      da : DATE := D#2021-05-07; db : DATE := D#2021-05-06; ta : TOD := TOD#10:00:00; tb : TOD := TOD#09:00:00;
      t23 : TOD := TOD#23:00:00; lx : LDT := LDT#2021-05-06-07:08:09; ly : LDT := LDT#2021-05-06-07:00:00;
      lh : LTIME := LT#1h; lh2 : LTIME := LT#2h; lt23 : LTOD := LTOD#23:00:00; lt12 : LTOD := LTOD#12:00:00;
      d20 : DATE := D#2020-01-01; one : INT := 1; two : INT := 2; three : INT := 3; four : INT := 4;
      y : INT := 2020; twelve : INT := 12; zero : INT; r15 : REAL := 1.5; tt : TIME := T#1h30m;
      sreal : STRING[8] := '1.5'; st : STRING[8] := 'T#5s'; sd : STRING[16] := 'D#2021-05-06'; sb : STRING[8] := 'TRUE';
      r16 : REAL := 16.0; r2 : REAL := 2.0; r100 : REAL := 100.0; l2r : LREAL := 2.0; l1e5 : LREAL := 1.0E5;
      ok : USINT; e1 : INT; hh, mm, ss, mss : INT;
  END_VAR
  VAR q AT %QB0 : USINT; q1 AT %QB1 : USINT; q2 AT %QB2 : USINT; q3 AT %QB3 : USINT; END_VAR
  ok := 0;
  IF d5 = dx + h THEN ok := ok + 1; END_IF;
  IF d6 = dx - h THEN ok := ok + 1; END_IF;
  IF t1 = dx - dy THEN ok := ok + 1; END_IF;
  IF t2 = da - db THEN ok := ok + 1; END_IF;
  IF t3 = t23 + h2 THEN ok := ok + 1; END_IF;
  IF t4 = ta - tb THEN ok := ok + 1; END_IF;
  IF l1 = lx + lh THEN ok := ok + 1; END_IF;
  IF l2 = lx - ly THEN ok := ok + 1; END_IF;
  IF l3 = CONCAT_LTOD(one, two, three, four) THEN ok := ok + 1; END_IF;
  IF l4 = CONCAT_LDT(y, one, one, twelve, zero, zero, zero) THEN ok := ok + 1; END_IF;
  IF l5 = CONCAT_DATE_LTOD(d20, lt12) THEN ok := ok + 1; END_IF;
  IF l6 = ADD_LTOD_LTIME(lt23, lh2) THEN ok := ok + 1; END_IF;
  IF s1 = REAL_TO_STRING(r15) THEN ok := ok + 1; END_IF;
  IF s3 = TIME_TO_STRING(tt) THEN ok := ok + 1; END_IF;
  IF s4 = DT_TO_STRING(dx) THEN ok := ok + 1; END_IF;
  IF r1 = STRING_TO_REAL(sreal) THEN ok := ok + 1; END_IF;
  IF tm = STRING_TO_TIME(st) THEN ok := ok + 1; END_IF;
  IF dd = STRING_TO_DATE(sd) THEN ok := ok + 1; END_IF;
  IF b1 = STRING_TO_BOOL(sb) THEN ok := ok + 1; END_IF;
  IF x1 = REAL_TO_INT(SQRT(r16)) THEN ok := ok + 1; END_IF;
  IF x3 = REAL_TO_INT(SQRT(r2) * r100) THEN ok := ok + 1; END_IF;
  IF x4 = 10.0 / SQRT(r2) THEN ok := ok + 1; END_IF;
  e1 := REAL_TO_INT(SQRT(r16));
  IF x5 = 100 / e1 THEN ok := ok + 1; END_IF;
  IF x11 = LREAL_TO_DINT(l1e5 * SQRT(l2r)) THEN ok := ok + 1; END_IF;
  q := ok;
  q1 := INT_TO_USINT(x1);
  q2 := INT_TO_USINT(x5);
  SPLIT_TOD(t3, hh, mm, ss, mss);
  q3 := INT_TO_USINT(hh);
END_PROGRAM
CONFIGURATION c RESOURCE r ON PLC TASK t(INTERVAL := T#10ms, PRIORITY := 1); PROGRAM p WITH t : main; END_RESOURCE END_CONFIGURATION

(* ---- control.st ---- *)
(* The ST statements: IF/ELSIF/ELSE, CASE with lists and ranges, FOR up
   and down with BY, WHILE, REPEAT, EXIT, RETURN. *)
PROGRAM main
VAR
  v AT %IW0 : INT;
  r_if AT %MW0 : INT;
  r_case AT %MW2 : INT;
  r_for AT %MD4 : DINT;
  r_down AT %MD8 : DINT;
  r_while AT %MW12 : INT;
  r_repeat AT %MW14 : INT;
  r_exit AT %MW16 : INT;
  r_ret AT %MW18 : INT;
END_VAR
VAR
  i : INT;
  j : INT;
END_VAR
IF v < 0 THEN
  r_if := -1;
ELSIF v = 0 THEN
  r_if := 0;
ELSIF v < 10 THEN
  r_if := 1;
ELSE
  r_if := 2;
END_IF;

CASE v OF
  0: r_case := 100;
  1, 2, 3: r_case := 200;
  4..9: r_case := 300 + v;
  -5..-1: r_case := -300;
ELSE
  r_case := 999;
END_CASE;

r_for := 0;
FOR i := 1 TO v BY 2 DO
  r_for := r_for + INT_TO_DINT(i);
END_FOR;
r_down := 0;
FOR i := 10 TO 1 BY -3 DO
  r_down := r_down * 10 + INT_TO_DINT(i);
END_FOR;

r_while := 0;
i := v;
WHILE i > 0 DO
  r_while := r_while + 1;
  i := i / 2;
END_WHILE;

r_repeat := 0;
REPEAT
  r_repeat := r_repeat + 1;
UNTIL r_repeat >= v
END_REPEAT;

r_exit := 0;
FOR i := 1 TO 10 DO
  FOR j := 1 TO 10 DO
    IF j > i THEN
      EXIT;
    END_IF;
    r_exit := r_exit + 1;
  END_FOR;
  IF i >= v THEN
    EXIT;
  END_IF;
END_FOR;

r_ret := 1;
IF v = 7 THEN
  RETURN;
END_IF;
r_ret := 2;
END_PROGRAM

CONFIGURATION plant
  RESOURCE r ON PLC
    TASK fast(INTERVAL := T#10ms, PRIORITY := 0);
    PROGRAM p WITH fast : main;
  END_RESOURCE
END_CONFIGURATION

(* ---- convert.st ---- *)
(* Conversions to and from STRING where the reference compiler's text and iecf's agree
   (docs/dependencies.md): integers in decimal, BOOL as TRUE and FALSE,
   a REAL whose shortest text is its %g, and reading them back - a
   number from the inputs there and back again. The rest of the text,
   which the reference compiler writes otherwise (a REAL's 10 digits, 16#ff for a bit
   string, every unit of a TIME), is runtime/tests/strings.c's. *)
PROGRAM main
VAR
  a AT %IW0 : INT;
  b AT %ID2 : DINT;
  r_back AT %MW0 : INT;
  r_len AT %MW2 : INT;
  r_dint AT %MD4 : DINT;
  r_real AT %MD8 : REAL;
  r_cmp AT %MW12 : WORD;
END_VAR
VAR
  text : STRING;
END_VAR
text := INT_TO_STRING(a);
r_len := LEN(text);
r_back := STRING_TO_INT(text) / 2;
r_dint := STRING_TO_DINT(CONCAT(DINT_TO_STRING(b), '0'));
r_real := STRING_TO_REAL(REAL_TO_STRING(INT_TO_REAL(a) / 4.0)) * 2.0;
r_cmp := 0;
IF BOOL_TO_STRING(a > 0) = 'TRUE' THEN r_cmp := r_cmp OR 1; END_IF;
IF BOOL_TO_STRING(a > 0) = 'FALSE' THEN r_cmp := r_cmp OR 2; END_IF;
IF REAL_TO_STRING(INT_TO_REAL(a) / 4.0) = '2.5' THEN r_cmp := r_cmp OR 4; END_IF;
IF STRING_TO_BOOL('TRUE') THEN r_cmp := r_cmp OR 8; END_IF;
IF DINT_TO_STRING(b) = '-123456' THEN r_cmp := r_cmp OR 16; END_IF;
END_PROGRAM

CONFIGURATION config
  RESOURCE res ON PLC
    TASK t(INTERVAL := T#10ms, PRIORITY := 0);
    PROGRAM p WITH t : main;
  END_RESOURCE
END_CONFIGURATION

(* ---- dates.st ---- *)
(* DATE, TOD and DT (Ed.3 Table 35; docs/dependencies.md): a TOD and a DT
   go on 7 hours a tick, from TOD#20:00:00 and DT#2026-11-07-22:00:00; each
   tick shows, as bits, comparisons of what Table 35's operators and
   functions give (DAY_OF_WEEK, which the reference compiler lacks, is
   runtime/tests/dates.c's). A TOD wraps at midnight in
   iecf, where the reference compiler's goes on past 24 hours: at tick 0 the TOD is
   TOD#03:00:00 in iecf and 27 hours in the reference compiler. iecf's trace is
   dates.iecf.trace. *)
PROGRAM main
VAR
  r_bits AT %MW0 : WORD;
END_VAR
VAR
  clock : TOD := TOD#20:00:00;
  stamp : DT := DT#2026-11-07-22:00:00;
  day : DATE;
  start : DT := DT#2026-11-07-00:00:00;
END_VAR
clock := clock + T#7h;
stamp := ADD_DT_TIME(stamp, T#7h);
day := DT_TO_DATE(stamp);
r_bits := 0;
IF clock < TOD#12:00:00 THEN r_bits := r_bits OR 16#0001; END_IF;
IF stamp > DT#2026-11-08-12:00:00 THEN r_bits := r_bits OR 16#0002; END_IF;
IF stamp - start > T#1d THEN r_bits := r_bits OR 16#0004; END_IF;
IF DT_TO_TOD(stamp) - clock = T#2h THEN r_bits := r_bits OR 16#0008; END_IF;
IF CONCAT_DATE_TOD(day, DT_TO_TOD(stamp)) = stamp THEN r_bits := r_bits OR 16#0010; END_IF;
IF SUB_DATE_DATE(day, D#2026-11-07) >= T#1d THEN r_bits := r_bits OR 16#0020; END_IF;
IF day = D#2026-11-09 THEN r_bits := r_bits OR 16#0040; END_IF;
IF SUB_DT_TIME(stamp, T#1d) < start THEN r_bits := r_bits OR 16#0080; END_IF;
IF clock - T#21h = TOD#06:00:00 THEN r_bits := r_bits OR 16#0100; END_IF;
IF SUB_TOD_TOD(TOD#01:00:00, TOD#23:00:00) = T#-22h THEN r_bits := r_bits OR 16#0200; END_IF;
IF MAX(clock, TOD#10:00:00) = clock THEN r_bits := r_bits OR 16#0400; END_IF;
IF DT_TO_DATE(DT#2026-11-07-23:59:59) = D#2026-11-07 THEN r_bits := r_bits OR 16#0800; END_IF;
END_PROGRAM

CONFIGURATION plant
  RESOURCE r ON PLC
    TASK fast(INTERVAL := T#10ms, PRIORITY := 0);
    PROGRAM p WITH fast : main;
  END_RESOURCE
END_CONFIGURATION

(* ---- durations.st ---- *)
(* A duration times or divided by a number (Ed.3 Table 35: MUL_TIME,
   DIV_TIME, * and /): by an integer exact, by a REAL rounded to whole
   milliseconds half to even, as REAL_TO_DINT rounds (docs/dependencies.md).
   The factor n comes from %IW0, 1 to 4 over the ticks; each bit is a
   comparison. iecf's TIME counts whole milliseconds (dividing like DINT,
   toward 0); the reference compiler's holds nanoseconds, so its T#10s / 3 is
   3.333333333s, T#3ms * 1.5 is 4.5ms and T#-7ms / 2 is -3.5ms, none
   equal to the whole milliseconds they are compared with: iecf's trace
   is durations.iecf.trace. LTIME, which
   the reference compiler lacks, MUL_TIME and DIV_TIME (the reference compiler has Ed.2's MULTIME and
   DIVTIME) and a number times a duration, n * T#1s (the reference compiler's C passes
   __time_mul its arguments the wrong way round and does not compile),
   are the generator's tests'. *)
PROGRAM main
VAR
  n AT %IW0 : INT;
  r_bits AT %MW0 : WORD;
END_VAR
VAR
  t : TIME;
  f : REAL;
END_VAR
r_bits := 0;
t := T#1s500ms * n;
IF t = T#1500ms * INT_TO_DINT(n) AND t > T#1s THEN r_bits := r_bits OR 16#0001; END_IF;
IF T#250ms * n = T#1s THEN r_bits := r_bits OR 16#0002; END_IF;
IF T#1s / n = T#250ms THEN r_bits := r_bits OR 16#0004; END_IF;
IF T#10s / n = T#3s333ms THEN r_bits := r_bits OR 16#0008; END_IF;
f := INT_TO_REAL(n) / 2.0;
IF T#1s * f = T#2s THEN r_bits := r_bits OR 16#0010; END_IF;
IF T#3ms * f = T#4ms THEN r_bits := r_bits OR 16#0020; END_IF;
IF MUL(T#100ms, n) = T#300ms THEN r_bits := r_bits OR 16#0040; END_IF;
IF DIV(T#1m, n) = T#20s THEN r_bits := r_bits OR 16#0080; END_IF;
IF T#1s / f = T#500ms THEN r_bits := r_bits OR 16#0100; END_IF;
IF T#-7ms / n = T#-3ms THEN r_bits := r_bits OR 16#0200; END_IF;
END_PROGRAM

CONFIGURATION plant
  RESOURCE r ON PLC
    TASK fast(INTERVAL := T#10ms, PRIORITY := 0);
    PROGRAM p WITH fast : main;
  END_RESOURCE
END_CONFIGURATION

(* ---- dynmem.st ---- *)
(* __NEW and __DELETE (the dynamic-memory extension), from the task's
   pool of 4096 bytes. Worked by hand: each tick a block one INT longer
   is taken, the list copied into it, its last element (count + 1) * 10,
   the old list given back: %QB0 the count, %QB1 the sum / 10 - tick 0:
   1 and 1, tick 1: 2 and 3, tick 2: 3 and 6, tick 3: 4 and 10. A pair
   from __NEW has its initial value, x 5 (%QB2), and __DELETE sets pr to
   0 (%QB3 1); 100000 INTs fit no pool of 4096 bytes: 0 (%QB4 1). At
   tick 3 a copy of a block given back is read: IECF_FAULT_NULL on line
   47, %QB5 left at 7.
   reference-skip: __NEW and __DELETE are CODESYS's, not IEC 61131-3. *)
TYPE pair : STRUCT x : INT := 5; y : INT; END_STRUCT; END_TYPE
PROGRAM main
  VAR
    list, grown, big, stale, copy : POINTER TO INT;
    pr : POINTER TO pair;
    count, i, sum : INT;
  END_VAR
  VAR q0 AT %QB0 : SINT; q1 AT %QB1 : SINT; q2 AT %QB2 : SINT; q3 AT %QB3 : SINT; q4 AT %QB4 : SINT;
      q5 AT %QB5 : SINT; END_VAR
  grown := __NEW(INT, count + 1);
  FOR i := 0 TO count - 1 DO
    grown[i] := list[i];
  END_FOR;
  grown[count] := (count + 1) * 10;
  IF list <> 0 THEN
    __DELETE(list);
  END_IF;
  list := grown;
  count := count + 1;
  sum := 0;
  FOR i := 0 TO count - 1 DO
    sum := sum + list[i];
  END_FOR;
  q0 := INT_TO_SINT(count);
  q1 := INT_TO_SINT(sum / 10);
  pr := __NEW(pair);
  q2 := INT_TO_SINT(pr^.x);
  __DELETE(pr);
  q3 := BOOL_TO_SINT(pr = 0);
  big := __NEW(INT, 100000);
  q4 := BOOL_TO_SINT(big = 0);
  IF count = 4 THEN
    stale := __NEW(INT, 2);
    copy := stale;
    __DELETE(stale);
    q5 := 7;
    q5 := INT_TO_SINT(copy[0]);
  END_IF;
END_PROGRAM

CONFIGURATION cf
  RESOURCE r ON x
    TASK tk(INTERVAL := T#10ms, PRIORITY := 1);
    PROGRAM p WITH tk : main;
  END_RESOURCE
END_CONFIGURATION

(* ---- edges.st ---- *)
(* The counters and bistables of Ed.3 Tables 43-45: CTU, CTD, CTUD, R_TRIG,
   F_TRIG, SR and RS.

   The reference compiler's counters stop where Ed.3 Table 45 does not: CTU and CTUD count
   up only while CV < PV, and CTD down only while CV > 0, where the table
   has CV < PVmax and CV > PVmin (each implementer-specific). Four CU
   pulses against a PV of 3 show it: the reference compiler's CTU stops at 3 and its CTUD
   at its loaded 2. iecf counts over the type's whole range, as decided
   (docs/dependencies.md): CTU to 4, CTUD to 6, and CTUD below 0 at the
   last CD. Its trace is edges.iecf.trace. *)
PROGRAM main
VAR
  cu AT %IX0.0 : BOOL;
  cd AT %IX0.1 : BOOL;
  rst AT %IX0.2 : BOOL;
  ld AT %IX0.3 : BOOL;
  s1 AT %IX0.4 : BOOL;
  r1 AT %IX0.5 : BOOL;
  up_q AT %QX0.0 : BOOL;
  dn_q AT %QX0.1 : BOOL;
  ud_qu AT %QX0.2 : BOOL;
  ud_qd AT %QX0.3 : BOOL;
  rise AT %QX0.4 : BOOL;
  fall AT %QX0.5 : BOOL;
  sr_q AT %QX0.6 : BOOL;
  rs_q AT %QX0.7 : BOOL;
  up_cv AT %MW0 : INT;
  dn_cv AT %MW2 : INT;
  ud_cv AT %MW4 : INT;
END_VAR
VAR
  c_up : CTU;
  c_dn : CTD;
  c_ud : CTUD;
  e_r : R_TRIG;
  e_f : F_TRIG;
  b_sr : SR;
  b_rs : RS;
END_VAR
c_up(CU := cu, R := rst, PV := 3);
c_dn(CD := cd, LD := ld, PV := 2);
c_ud(CU := cu, CD := cd, R := rst, LD := ld, PV := 2);
e_r(CLK := cu);
e_f(CLK := cu);
b_sr(S1 := s1, R := r1);
b_rs(S := s1, R1 := r1);
up_q := c_up.Q;
up_cv := c_up.CV;
dn_q := c_dn.Q;
dn_cv := c_dn.CV;
ud_qu := c_ud.QU;
ud_qd := c_ud.QD;
ud_cv := c_ud.CV;
rise := e_r.Q;
fall := e_f.Q;
sr_q := b_sr.Q1;
rs_q := b_rs.Q1;
END_PROGRAM

CONFIGURATION plant
  RESOURCE r ON PLC
    TASK fast(INTERVAL := T#10ms, PRIORITY := 0);
    PROGRAM p WITH fast : main;
  END_RESOURCE
END_CONFIGURATION

(* ---- enable.st ---- *)
(* EN and ENO on a call (Ed.3 6.6.1.5; docs/behaviour/en-eno.md): with
   EN FALSE the call does not happen and its statement is left undone,
   the target keeping its value; ENO is FALSE then, and when the
   function's own operation flags. %IX0.0 is EN over the ticks; the
   divisor %IW2 is 0 at tick 2, when EN is FALSE, so DIV is not called
   and nothing faults. The reference compiler, by its own reading, assigns the function's
   default result when EN is FALSE, and keeps ENO TRUE through an
   overflow: iecf's trace is enable.iecf.trace. *)
FUNCTION twice : INT
VAR_INPUT x : INT; END_VAR
twice := x * 2;
END_FUNCTION

PROGRAM main
VAR
  go AT %IX0.0 : BOOL;
  d AT %IW2 : INT;
  r_div AT %MW0 : INT;
  r_twice AT %MW2 : INT;
  r_eno AT %MB4 : BYTE;
END_VAR
VAR
  ok1, ok2, ok3 : BOOL;
  n : INT := 16000;
END_VAR
r_div := DIV(EN := go, IN1 := INT#100, IN2 := d, ENO => ok1);
r_twice := twice(EN := go, x := n, ENO => ok2);
n := n + 100;
r_eno := 0;
IF ok1 THEN r_eno := r_eno OR 1; END_IF;
IF ok2 THEN r_eno := r_eno OR 2; END_IF;
END_PROGRAM

CONFIGURATION plant
  RESOURCE res ON PLC
    TASK fast(INTERVAL := T#10ms, PRIORITY := 0);
    PROGRAM p WITH fast : main;
  END_RESOURCE
END_CONFIGURATION

(* ---- extcompare.st ---- *)
(* GT, GE, EQ, LE and LT with more than two inputs (Ed.3 Table 33:
   each neighbouring pair holds), every input computed once and in
   order; the negation of a TIME and an LTIME; the shifts and rotations
   of a BOOL. Worked by hand, the same at every tick:
   v 5: GT(v, 2, 1) TRUE (%QX0.0); GT(v, 6, 1) FALSE (%QX0.1);
   GE(v, 5, 5, 1) TRUE (%QX0.2); LT(1, 2, 2) FALSE (%QX0.3);
   LE(1, 2, 2) TRUE (%QX0.4). s 'ab': EQ('ab', s, 'ab') TRUE (%QX0.5).
   t T#2s: LT(T#1s, t, T#3s) TRUE (%QX0.6).
   Inc adds 1 to its in-out and gives it. n := 0; GT(10, Inc(n), 0):
   Inc is called once, n is 1 (%QB1), and 10 > 1 > 0 TRUE (%QX0.7).
   GT(n, Inc(n), 0): n is read first, 1, then Inc makes it 2: 1 > 2 is
   FALSE (%QX2.0), and n is 2 (%QB3).
   -T#1s500ms is T#-1s500ms (%QX2.1); -LTIME#2ns is LTIME#-2ns
   (%QX2.2). A BOOL is one bit: SHL(TRUE, 0) TRUE (%QX2.3), SHL(TRUE,
   1) FALSE (%QX2.4), ROL(TRUE, 5) TRUE (%QX2.5), SHR(TRUE, 1) FALSE
   (%QX2.6), ROR(TRUE, 2) TRUE (%QX2.7).
   Last, the TIME DINT's lowest, T#-24d20h31m23s648ms, negated: it
   wraps to itself and is flagged OVERFLOW (%QB4 1).
   reference-skip: no LTIME; -t on a TIME and SHL on a BOOL: its C
   does not build. *)
FUNCTION Inc : INT
  VAR_IN_OUT io : INT; END_VAR
  io := io + 1;
  Inc := io;
END_FUNCTION
PROGRAM main
  VAR
    v : INT := 5;
    n : INT;
    s : STRING := 'ab';
    t : TIME := T#2s;
    t2 : TIME;
    l2 : LTIME;
    bb : BOOL := TRUE;
    tm : TIME;
  END_VAR
  VAR
    q00 AT %QX0.0 : BOOL;
    q01 AT %QX0.1 : BOOL;
    q02 AT %QX0.2 : BOOL;
    q03 AT %QX0.3 : BOOL;
    q04 AT %QX0.4 : BOOL;
    q05 AT %QX0.5 : BOOL;
    q06 AT %QX0.6 : BOOL;
    q07 AT %QX0.7 : BOOL;
    q1 AT %QB1 : SINT;
    q20 AT %QX2.0 : BOOL;
    q21 AT %QX2.1 : BOOL;
    q22 AT %QX2.2 : BOOL;
    q23 AT %QX2.3 : BOOL;
    q24 AT %QX2.4 : BOOL;
    q25 AT %QX2.5 : BOOL;
    q26 AT %QX2.6 : BOOL;
    q27 AT %QX2.7 : BOOL;
    q3 AT %QB3 : SINT;
    q4 AT %QB4 : SINT;
  END_VAR
  q00 := GT(v, 2, 1);
  q01 := GT(v, 6, 1);
  q02 := GE(v, 5, 5, 1);
  q03 := LT(1, 2, 2);
  q04 := LE(1, 2, 2);
  q05 := EQ('ab', s, 'ab');
  q06 := LT(T#1s, t, T#3s);
  n := 0;
  q07 := GT(10, Inc(n), 0);
  q1 := INT_TO_SINT(n);
  q20 := GT(n, Inc(n), 0);
  q3 := INT_TO_SINT(n);
  t2 := T#1s500ms;
  t2 := -t2;
  q21 := t2 = T#-1s500ms;
  l2 := LTIME#2ns;
  l2 := -l2;
  q22 := l2 = LTIME#-2ns;
  q23 := SHL(bb, 0);
  q24 := SHL(bb, 1);
  q25 := ROL(bb, 5);
  q26 := SHR(bb, 1);
  q27 := ROR(bb, 2);
  tm := T#-24d20h31m23s648ms;
  tm := -tm;
  IF tm = T#-24d20h31m23s648ms THEN
    q4 := 1;
  END_IF;
END_PROGRAM

CONFIGURATION c
  RESOURCE r ON x
    TASK t(INTERVAL := T#10ms, PRIORITY := 1);
    PROGRAM p WITH t : main;
  END_RESOURCE
END_CONFIGURATION

(* ---- flexcopy.st ---- *)
(* A whole ARRAY[*] assigned (Ed.3 6.5.3; docs/dependencies.md): from
   another ARRAY[*] or from an array of fixed bounds, of as many
   elements in each dimension - which only the run knows, so it is
   checked as the assignment runs: a fault (index) and nothing copied
   when they differ. The bounds themselves need not match.
   COPY does dst := src. FILL3 does dst := three, its own [7, 8, 9].
   GRID does dst := src for two dimensions.
   Worked by hand, k %IB0 1, 2, 3:
   a: 1..3, [1, 2, 3]; b: -1..1, [0, 0, 0]. COPY(b, a) at tick 0: b
   [1, 2, 3]: b[-1] 1 (%QB0), b[1] 3 (%QB1).
   FILL3(a): a [7, 8, 9]: a[2] 8 (%QB2); then a[1] := k. So at the
   ticks after the first, COPY(b, a) gives b [k of the tick before, 8,
   9]: %QB0 1, 1, 2 and %QB1 3, 9, 9.
   m: 1..2, 0..1, [[1, 2], [3, 4]]; n: 0..1, 5..6. GRID(n, m): n[1, 6]
   4 (%QB3).
   Onto itself: COPY(a, a) leaves a as it is: a[3] 9 (%QB4).
   At tick 2, COPY(w, a) with w of 2 elements: 2 is not 3, a fault
   (index) in COPY at its assignment; w is as it was, w[1] 0 (%QB5),
   read before the call.
   reference-skip: ARRAY[*] is Ed.3's; the reference compiler (Ed.2)
   has none. *)
FUNCTION COPY
  VAR_IN_OUT dst, src : ARRAY [*] OF INT; END_VAR
  dst := src;
END_FUNCTION
FUNCTION FILL3
  VAR_IN_OUT dst : ARRAY [*] OF INT; END_VAR
  VAR three : ARRAY [1..3] OF INT := [7, 8, 9]; END_VAR
  dst := three;
END_FUNCTION
FUNCTION GRID
  VAR_IN_OUT dst, src : ARRAY [*, *] OF INT; END_VAR
  dst := src;
END_FUNCTION
CONFIGURATION c
  RESOURCE r ON PLC
    TASK t(INTERVAL := T#10ms, PRIORITY := 1);
    PROGRAM p WITH t : main;
  END_RESOURCE
END_CONFIGURATION
PROGRAM main
  VAR
    a : ARRAY [1..3] OF INT := [1, 2, 3];
    b : ARRAY [-1..1] OF INT;
    m : ARRAY [1..2, 0..1] OF INT := [1, 2, 3, 4];
    n : ARRAY [0..1, 5..6] OF INT;
    w : ARRAY [0..1] OF INT;
  END_VAR
  VAR k AT %IB0 : SINT; END_VAR
  VAR
    q0 AT %QB0 : SINT;
    q1 AT %QB1 : SINT;
    q2 AT %QB2 : SINT;
    q3 AT %QB3 : SINT;
    q4 AT %QB4 : SINT;
    q5 AT %QB5 : SINT;
  END_VAR
  COPY(b, a);
  q0 := INT_TO_SINT(b[-1]);
  q1 := INT_TO_SINT(b[1]);
  FILL3(a);
  q2 := INT_TO_SINT(a[2]);
  a[1] := k;
  GRID(n, m);
  q3 := INT_TO_SINT(n[1, 6]);
  COPY(a, a);
  q4 := INT_TO_SINT(a[3]);
  q5 := INT_TO_SINT(w[1]);
  IF k = 3 THEN
    COPY(w, a);
  END_IF;
END_PROGRAM

(* ---- fneffen.st ---- *)
(* EN on a call of a FUNCTION with effects (Ed.3 6.6.1.5): an in-out and
   an output (bump), a VAR_EXTERNAL written (tick), no result (addw).
   EN FALSE: the function is not called - its in-outs, outputs and
   globals are left as they were - ENO is FALSE, and the statement is
   left undone; ENO is FALSE too when the call's own operation raised a
   flag; not when storing its outputs does (an output clamped into a
   subrange).
   Worked by hand, v 0, r -1, t -1, w 32766, g 0 at the start:
   u 0, s 0:
   Tick 0, run TRUE: bump: v 2, t 4, r 2; tick: g 1, qg 1; addw: w 32767,
   qok TRUE; bump: u 2, s 4, qok2 TRUE.
   Tick 1, run FALSE: nothing called: v 2, r 2, t 4, qg 1, w 32767, u 2,
   s 4; qok, qok2 FALSE.
   Tick 2, run TRUE: v 4, t 8, r 4; g 2, qg 2; addw: w 32767 + 1 wraps to
   -32768, flag OVERFLOW in addw on line 39, qok FALSE; bump: u 4, its
   output 8 clamped to s 5 (flagged too, after the first), qok2 TRUE.
   reference-skip: the reference compiler (Ed.2) refuses VAR_EXTERNAL in
   a FUNCTION. *)
TYPE small : INT (0..5); END_TYPE

FUNCTION bump : INT
VAR_IN_OUT x : INT; END_VAR
VAR_INPUT d : INT; END_VAR
VAR_OUTPUT twice : INT; END_VAR
x := x + d;
twice := x * 2;
bump := x;
END_FUNCTION

FUNCTION tick : INT
VAR_EXTERNAL g : INT; END_VAR
g := g + 1;
tick := g;
END_FUNCTION

FUNCTION addw
VAR_IN_OUT x : INT; END_VAR
VAR_INPUT d : INT; END_VAR
x := x + d;
END_FUNCTION

PROGRAM main
VAR
  run AT %IX0.0 : BOOL;
  qv AT %QW0 : INT;
  qr AT %QW2 : INT;
  qt AT %QW4 : INT;
  qg AT %QW6 : INT;
  qok AT %QX8.0 : BOOL;
  qw AT %QW10 : INT;
  qok2 AT %QX8.1 : BOOL;
  qs AT %QW12 : INT;
END_VAR
VAR
  v : INT;
  r : INT := -1;
  t : INT := -1;
  w : INT := 32766;
  u, r2 : INT;
  s : small;
END_VAR
r := bump(EN := run, x := v, d := 2, twice => t);
qg := tick(EN := run);
addw(EN := run, x := w, d := 1, ENO => qok);
r2 := bump(EN := run, x := u, d := 2, twice => s, ENO => qok2);
qv := v;
qr := r;
qt := t;
qw := w;
qs := s;
END_PROGRAM

CONFIGURATION Plant
  VAR_GLOBAL g : INT; END_VAR
  RESOURCE r ON PLC
    TASK fast(INTERVAL := T#10ms, PRIORITY := 1);
    PROGRAM p WITH fast : main;
  END_RESOURCE
END_CONFIGURATION

(* ---- fninout.st ---- *)
(* A FUNCTION's in-outs (Ed.3 6.6.2.2, rule 6): an in-out reads and
   writes the variable the call passes, two at once in swap; an in-out
   passed on to another function's in-out, in twice. Externals are in
   fnorder: the reference compiler (Ed.2) refuses VAR_EXTERNAL in a
   FUNCTION. *)
FUNCTION swap : BOOL
VAR_IN_OUT a, b : INT; END_VAR
VAR t : INT; END_VAR
t := a;
a := b;
b := t;
swap := a > b;
END_FUNCTION

FUNCTION bump : INT
VAR_INPUT n : INT; END_VAR
VAR_IN_OUT v : INT; END_VAR
v := v + n * 3;
bump := v;
END_FUNCTION

FUNCTION twice : INT
VAR_IN_OUT w : INT; END_VAR
VAR k : INT; END_VAR
k := bump(n := 1, v := w);
twice := bump(n := 1, v := w);
END_FUNCTION

PROGRAM main
VAR
  vin AT %IW0 : INT;
  bin AT %IW2 : INT;
  qx AT %QW0 : INT;
  qy AT %QW2 : INT;
  qk AT %QW4 : INT;
  qok AT %QX6.0 : BOOL;
END_VAR
VAR
  x, y, k : INT;
  ok : BOOL;
END_VAR
x := vin;
y := bin;
ok := swap(a := x, b := y);
qok := ok;
k := bump(n := 2, v := x);
k := twice(w := y);
qx := x;
qy := y;
qk := k;
END_PROGRAM

CONFIGURATION Plant
  RESOURCE r ON PLC
    TASK fast(INTERVAL := T#10ms, PRIORITY := 1);
    PROGRAM p WITH fast : main;
  END_RESOURCE
END_CONFIGURATION

(* ---- fnorder.st ---- *)
(* A FUNCTION's externals (Ed.3 6.6.2.2, rules 4-5), and the order of
   evaluation once a call has effects (7.3.2, rule 3: "the leftmost
   operand shall be evaluated first"):
   - x + bump(1, x): x read before the call changes it;
   - bump(1, y) * 10 + y: y read after it;
   - bump(1, w) - bump(2, w): the left call first;
   - peek() + bump(1, w) + peek(): total read, written, read again;
   - x + mark(q => x): x read before the call's output is stored in it;
   - 100 / zin + mark(q => qm): the division first, so at tick 1, zin 0,
     it faults before mark runs, and qm, cleared just before, stays 0.
   An in-out given an element by a computed index, arr[i].
   Worked by hand: tick 0, vin 2, zin 1: qa 7, qb 55, qc -6, qd 15,
   qt 11, qp 23 (5 + 12 + 6), qe 101, qm 1. Tick 1, vin -3, zin 0: qa -3,
   qb 0, qc -6, qd 15, qt 22, qp 45 (16 + 12 + 17), qe 101, qm 0, fault
   DIVISION_BY_ZERO; total grows by every bump's n, 11 a tick. qf is
   vin + 1: 3, then -2.
   reference-skip: the reference compiler (Ed.2) refuses VAR_EXTERNAL in
   a FUNCTION. *)
FUNCTION bump : INT
VAR_INPUT n : INT; END_VAR
VAR_IN_OUT v : INT; END_VAR
VAR_EXTERNAL total : DINT; END_VAR
VAR_EXTERNAL CONSTANT k3 : INT; END_VAR
v := v + n * k3;
total := total + n;
bump := v;
END_FUNCTION

FUNCTION peek : DINT
VAR_EXTERNAL total : DINT; END_VAR
peek := total;
END_FUNCTION

FUNCTION mark : INT
VAR_OUTPUT q : INT; END_VAR
q := 1;
mark := 1;
END_FUNCTION

PROGRAM main
VAR
  vin AT %IW0 : INT;
  zin AT %IW2 : INT;
  qa AT %QW0 : INT;
  qb AT %QW2 : INT;
  qc AT %QW4 : INT;
  qd AT %QW6 : INT;
  qt AT %QD8 : DINT;
  qp AT %QD12 : DINT;
  qe AT %QW16 : INT;
  qm AT %QW18 : INT;
  qf AT %QW20 : INT;
END_VAR
VAR
  x, y, w, i : INT;
  arr : ARRAY[0..3] OF INT;
END_VAR
VAR_EXTERNAL total : DINT; END_VAR
x := vin;
qa := x + bump(1, x);
y := vin;
qb := bump(1, y) * 10 + y;
w := 0;
qc := bump(1, w) - bump(2, w);
qp := peek() + bump(1, w) + peek();
i := vin MOD 4;
IF i < 0 THEN i := 0; END_IF;
qd := bump(5, arr[i]);
qt := total;
x := vin;
qf := x + mark(q => x);
qm := 0;
qe := 100 / zin + mark(q => qm);
END_PROGRAM

CONFIGURATION Plant
  VAR_GLOBAL
    total : DINT;
  END_VAR
  VAR_GLOBAL CONSTANT
    k3 : INT := 3;
  END_VAR
  RESOURCE r ON PLC
    TASK fast(INTERVAL := T#10ms, PRIORITY := 1);
    PROGRAM p WITH fast : main;
  END_RESOURCE
END_CONFIGURATION

(* ---- fnout.st ---- *)
(* A FUNCTION's outputs (Ed.3 6.6.1.4, 6.6.2.2): taken with =>, into a
   variable and a variable at an address; set from the call, an output's initial value at each call, as
   a FUNCTION has no memory; RETURN gives the outputs as they are.
   divmod(5, 0) returns before it sets q and r: q 0, r its initial -1.
   count's output starts at 0 at each call, so it always gives 1. An
   output into an array element is in fnoutx: the reference compiler's
   C for it does not compile. *)
FUNCTION divmod : INT
VAR_INPUT a, b : INT; END_VAR
VAR_OUTPUT q : INT; r : INT := -1; END_VAR
IF b = 0 THEN RETURN; END_IF;
q := a / b;
r := a MOD b;
divmod := 1;
END_FUNCTION

FUNCTION count : INT
VAR_OUTPUT n : INT; END_VAR
n := n + 1;
count := n;
END_FUNCTION

PROGRAM main
VAR
  vin AT %IW0 : INT;
  bin AT %IW2 : INT;
  qq AT %QW0 : INT;
  qr AT %QW2 : INT;
  qk AT %QW4 : INT;
  qn AT %QW6 : INT;
  qa AT %QW8 : INT;
END_VAR
VAR
  k, n, m : INT;
END_VAR
qk := divmod(a := vin, b := bin, q => qq, r => qr);
k := count(n => n);
qk := qk + k * 10;
qn := n;
k := divmod(a := 9, b := 4, r => m);
qa := m + k * 10;
END_PROGRAM

CONFIGURATION Plant
  RESOURCE r ON PLC
    TASK fast(INTERVAL := T#10ms, PRIORITY := 1);
    PROGRAM p WITH fast : main;
  END_RESOURCE
END_CONFIGURATION

(* ---- fnoutx.st ---- *)
(* A FUNCTION's outputs as the reference compiler does not take them:
   negated (NOT neg =>), widened into a DINT and a LINT (Ed.3 6.6.1.6,
   rule 5), given in order where declared, all of them (Ed.3
   6.6.1.4.2: divmod(vin, 4, ql, dr, dn)), into an array element by a
   computed index; and a call that faults: divmod(1, 0)
   divides by zero, the task stops, and nothing is stored - its output
   and its result are both for qs, which keeps the 5 it was just given.
   An output is stored before the statement's own target: qs := divmod(
   ..., r => qs) leaves qs the result. split10 has no result (Ed.3
   6.6.2.1), called as a statement, in order: v, hi, lo, then the
   in-out calls, as declared.
   Worked by hand: tick 0, vin 7, bin 1: qd 2, ql 1, qp TRUE, arr[3] 2,
   qa 2000, qk 111, qs 1, qh 0, qlo 7, qn 1. Tick 1, vin -7, bin 0: qd -2, ql -1, qp FALSE,
   arr[0] 2, qa 2002, qk 111, qh 0, qlo -7, qn 2, qs 5, fault
   DIVISION_BY_ZERO in DIVMOD.
   reference-skip: the reference compiler crashes on NOT q =>, has no
   implicit conversions, its C for an output into an array element
   does not compile, and Ed.2 has no FUNCTION without a result. *)
FUNCTION divmod : INT
VAR_INPUT a, b : INT; END_VAR
VAR_OUTPUT q : INT; r : INT := -1; neg : BOOL; END_VAR
q := a / b;
r := a MOD b;
neg := q < 0;
divmod := 1;
END_FUNCTION

FUNCTION split10
VAR_INPUT v : INT; END_VAR
VAR_OUTPUT hi, lo : INT; END_VAR
VAR_IN_OUT calls : INT; END_VAR
hi := v / 10;
lo := v MOD 10;
calls := calls + 1;
END_FUNCTION

PROGRAM main
VAR
  vin AT %IW0 : INT;
  bin AT %IW2 : INT;
  qd AT %QD0 : DINT;
  ql AT %QL4 : LINT;
  qp AT %QX12.0 : BOOL;
  qa AT %QW14 : INT;
  qk AT %QW16 : INT;
  qs AT %QW18 : INT;
  qh AT %QW20 : INT;
  qlo AT %QW22 : INT;
  qn AT %QW24 : INT;
END_VAR
VAR
  i, n, dr : INT;
  dn : BOOL;
  arr : ARRAY[0..3] OF INT;
END_VAR
qk := divmod(a := vin, b := 3, q => qd, NOT neg => qp);
qk := qk + divmod(vin, 4, ql, dr, dn) * 10;
i := vin MOD 4;
IF i < 0 THEN i := 0; END_IF;
qk := qk + divmod(a := 9, b := 4, q => arr[i]) * 100;
qa := arr[0] + arr[1] * 10 + arr[2] * 100 + arr[3] * 1000;
split10(vin, qh, qlo, n);
qn := n;
qs := 5;
qs := divmod(a := 1, b := bin, r => qs);
END_PROGRAM

CONFIGURATION Plant
  RESOURCE r ON PLC
    TASK fast(INTERVAL := T#10ms, PRIORITY := 1);
    PROGRAM p WITH fast : main;
  END_RESOURCE
END_CONFIGURATION

(* ---- functions.st ---- *)
(* The operators as functions (Ed.3 Tables 29-31, 33): ADD, MUL, AND,
   OR, XOR with more than two inputs; SUB, DIV, MOD; NOT; the
   comparisons GT, GE, EQ, LE, LT, NE; MOVE; SEL; EXPT and **. These are
   what Prokop's ladder and function block diagrams are written in.
   EXPT's results here are exact in binary floating point. *)
PROGRAM main
VAR
  a AT %IW0 : INT;
  b AT %IW2 : INT;
  m AT %IB4 : BYTE;
  s AT %IX5.0 : BOOL;
  r_add AT %MW0 : INT;
  r_mul AT %MW2 : INT;
  r_sub AT %MW4 : INT;
  r_div AT %MW6 : INT;
  r_mod AT %MW8 : INT;
  r_and AT %MB10 : BYTE;
  r_or AT %MB11 : BYTE;
  r_xor AT %MB12 : BYTE;
  r_not AT %MB13 : BYTE;
  r_cmp AT %MB14 : BYTE;
  r_sel AT %MW16 : INT;
  r_move AT %MW18 : INT;
  r_expt AT %MD20 : REAL;
  r_pow AT %ML24 : LREAL;
  r_bool AT %QX0.0 : BOOL;
END_VAR
r_add := ADD(a, b, 3);
r_mul := MUL(a, 2, -1);
r_sub := SUB(a, b);
r_div := DIV(a, b);
r_mod := MOD(a, b);
r_and := AND(m, BYTE#16#F0, BYTE#16#3C);
r_or := OR(m, BYTE#16#01);
r_xor := XOR(m, BYTE#16#FF, BYTE#16#0F);
r_not := NOT(m);
r_cmp := 0;
IF GT(a, b) THEN r_cmp := r_cmp OR 1; END_IF;
IF GE(a, b) THEN r_cmp := r_cmp OR 2; END_IF;
IF EQ(a, b) THEN r_cmp := r_cmp OR 4; END_IF;
IF LE(a, b) THEN r_cmp := r_cmp OR 8; END_IF;
IF LT(a, b) THEN r_cmp := r_cmp OR 16; END_IF;
IF NE(a, b) THEN r_cmp := r_cmp OR 32; END_IF;
r_sel := SEL(s, a, b);
r_move := MOVE(b);
r_expt := EXPT(INT_TO_REAL(b), 2);
r_pow := INT_TO_LREAL(a) ** 2.0 + 2.0 ** b;
r_bool := AND(OR(s, r_bool), NOT(EQ(a, 0)));
END_PROGRAM

CONFIGURATION config
  RESOURCE res ON PLC
    TASK t(INTERVAL := T#10ms, PRIORITY := 0);
    PROGRAM p WITH t : main;
  END_RESOURCE
END_CONFIGURATION

(* ---- globalns.st ---- *)
(* The global-namespace extension (docs/extensions.md): `_.` names the
   global namespace (Siemens, PLCnext; NAMESPACES.md D4). Inside Plant,
   ABS is Plant's own, x + 1000, and _.ABS the standard one; Lib.twice
   is Plant.Lib's, 3 x, and _.Lib.twice the top-level Lib's, 2 x.
   Worked by hand, tick 0, vin -4: q0 = -4 + 1000 = 996; q1 = 4;
   q2 = -12; q3 = -8. Tick 1, vin 7: q0 1007; q1 7; q2 21; q3 14.
   reference-skip: an extension, and the reference compiler has no
   namespaces. *)
NAMESPACE Lib
    FUNCTION twice : INT
    VAR_INPUT x : INT; END_VAR
        twice := x * 2;
    END_FUNCTION
END_NAMESPACE

NAMESPACE Plant
    NAMESPACE Lib
        FUNCTION twice : INT
        VAR_INPUT x : INT; END_VAR
            twice := x * 3;
        END_FUNCTION
    END_NAMESPACE

    FUNCTION ABS : INT
    VAR_INPUT x : INT; END_VAR
        ABS := x + 1000;
    END_FUNCTION

    PROGRAM Main
    VAR
        vin AT %IW0 : INT;
        q0 AT %QW0 : INT;
        q1 AT %QW2 : INT;
        q2 AT %QW4 : INT;
        q3 AT %QW6 : INT;
    END_VAR
        q0 := ABS(vin);
        q1 := _.ABS(vin);
        q2 := Lib.twice(vin);
        q3 := _.Lib.twice(vin);
    END_PROGRAM
END_NAMESPACE

CONFIGURATION Works
  RESOURCE r ON PLC
    TASK fast(INTERVAL := T#10ms, PRIORITY := 1);
    PROGRAM p WITH fast : Plant.Main;
  END_RESOURCE
END_CONFIGURATION

(* ---- hierfault.st ---- *)
(* A hierarchical address the platform has not (docs/c-output.md §4):
   the harness's iecf_address gives NULL for a level of 99, so the start
   faults with IECF_FAULT_IMAGE before anything runs, and no task runs.
   hierfault.iecf.trace: the reference compiler takes the address as a
   variable of its own, with no platform to ask, so nothing faults. *)
PROGRAM main
  VAR x AT %IW99.1 : INT; END_VAR
  VAR q AT %QW0 : INT; END_VAR
  q := x + 1;
END_PROGRAM
CONFIGURATION c RESOURCE r ON PLC TASK t(INTERVAL := T#10ms, PRIORITY := 1); PROGRAM p WITH t : main; END_RESOURCE END_CONFIGURATION

(* ---- image.st ---- *)
(* The process image: each size of address, read and written; a located
   variable's initial value; %M as well as %Q. *)
PROGRAM main
VAR
  inp AT %IB0 : BYTE;
  bit AT %IX1.2 : BOOL;
  cnt AT %QW0 : INT;
  acc AT %QD2 : DINT := 100;
  flag AT %QX6.3 : BOOL;
  big AT %ML0 : LINT;
  w AT %MW8 : WORD := 16#ABCD;
END_VAR
cnt := cnt + BYTE_TO_INT(inp);
acc := acc - 7;
flag := bit;
big := big + LINT#4294967296;
w := ROL(w, 4);
END_PROGRAM

CONFIGURATION plant
  RESOURCE r ON PLC
    TASK fast(INTERVAL := T#10ms, PRIORITY := 0);
    PROGRAM p WITH fast : main;
  END_RESOURCE
END_CONFIGURATION

(* ---- infinity.st ---- *)
(* An infinite or NaN REAL carries on and is flagged, not faulted
   (docs/c-output.md §5, decided 2026-11-06). At tick 1 the product
   overflows to +infinity; at tick 2 infinity minus infinity is a NaN.
   Both compilers write the same bytes and the program goes on counting;
   iecf's trace also shows ctx->flag: the first, an infinity (code 2) at
   line 21, stays until the platform clears it. *)
PROGRAM main
VAR
  k AT %IW0 : INT;
  r_mul AT %MD0 : REAL;
  r_diff AT %MD4 : REAL;
  ticks AT %MW8 : INT;
END_VAR
VAR
  x : REAL;
END_VAR
x := 1.0E5;
IF k >= 1 THEN
  x := 1.0E10;
END_IF;
r_mul := x * 1.0E30;
IF k >= 2 THEN
  r_diff := r_mul - r_mul;
END_IF;
ticks := ticks + 1;
END_PROGRAM

CONFIGURATION plant
  RESOURCE r ON PLC
    TASK fast(INTERVAL := T#10ms, PRIORITY := 0);
    PROGRAM p WITH fast : main;
  END_RESOURCE
END_CONFIGURATION

(* ---- initfault.st ---- *)
(* An initial value that faults as its variable is set up (the
   initial-expressions extension, docs/extensions.md): z is 0, so Quot(x,
   z) divides by zero in Quot, at its line (8). The fault stops the
   set-up there, as a statement's stops its body, and the program is
   stopped until the next start (docs/c-output.md §5): no task runs, and
   %QB0 stays 0.
   reference-skip: a variable in an initial value is not IEC 61131-3. *)
FUNCTION Quot : INT VAR_INPUT a, b : INT; END_VAR Quot := a / b; END_FUNCTION

PROGRAM main
  VAR
    z : INT;
    x : INT := 7;
    y : INT := Quot(x, z);
    w : INT := 3;
  END_VAR
  VAR q0 AT %QB0 : SINT; END_VAR
  q0 := INT_TO_SINT(x + y + w);
END_PROGRAM

CONFIGURATION c
  RESOURCE r ON x
    TASK t(INTERVAL := T#10ms, PRIORITY := 1);
    PROGRAM p WITH t : main;
  END_RESOURCE
END_CONFIGURATION

(* ---- inoutstop.st ---- *)
(* An element by an index out of bounds given to a FUNCTION's in-out
   of a structure: the statement stops before the call, which would
   have run on another element (docs/dependencies.md). fp writes g (Q1)
   when it runs: Q1 stays 00, Q0 is 07 from the line before, and the
   task faults (3, an index) at the call's line.
   reference-skip: VAR_IN_OUT of a FUNCTION, as `fnorder`. *)
TYPE pt : STRUCT x : INT; y : INT; END_STRUCT; END_TYPE
FUNCTION fp : INT
  VAR_IN_OUT p : pt; END_VAR
  VAR_EXTERNAL g : USINT; END_VAR
  g := 9;
  p.x := 1;
  fp := p.x;
END_FUNCTION
PROGRAM main
  VAR a : ARRAY [1..2] OF pt; k : INT := 3; r : INT; END_VAR
  VAR q AT %QB0 : USINT; END_VAR
  q := 7;
  r := fp(a[k]);
END_PROGRAM
CONFIGURATION c
  VAR_GLOBAL g AT %QB1 : USINT; END_VAR
  RESOURCE r ON PLC TASK t(INTERVAL := T#10ms, PRIORITY := 1); PROGRAM p WITH t : main; END_RESOURCE
END_CONFIGURATION

(* ---- intbits.st ---- *)
(* Three CODESYS ways with integers, each an extension. Worked by hand:
   integer-shifts: i := -8. SHR(i, 1) keeps the sign, -4 (%QW0);
   SHR(i, 20), past INT's 16 bits, -1 (%QW2); SHL(i, 2), -32 (%QW4);
   ROL(INT#-32768, 1), the top bit round to the bottom, 1 (%QW6);
   SHR(u, n) with UINT u 40000 and BYTE n 3, 5000 (%QW8).
   integer-bit-access: d := -2 (16#FFFFFFFE): d.0 FALSE, d.1 TRUE
   (%QX10.0, %QX10.1); d.0 := TRUE makes it -1 (%QD12); k := 5, k.%X15 :=
   TRUE sets INT's sign bit, -32763 (%QW16).
   integer-expt: EXPT(2, n) with INT n 10, 1024.0 as REAL, 1024 (%QW18);
   EXPT(q, 3) with DINT q -3, an LREAL, -27.0, -27 (%QW20).
   reference-skip: none of the three is IEC 61131-3. *)
PROGRAM main
  VAR
    i : INT := -8; u : UINT := 40000; n : BYTE := 3; d : DINT := -2; k : INT := 5;
    e : INT := 10; base : INT := 2; q : DINT := -3;
  END_VAR
  VAR
    q0 AT %QW0 : INT; q1 AT %QW2 : INT; q2 AT %QW4 : INT; q3 AT %QW6 : INT; q4 AT %QW8 : UINT;
    b0 AT %QX10.0 : BOOL; b1 AT %QX10.1 : BOOL; q5 AT %QD12 : DINT; q6 AT %QW16 : INT;
    q7 AT %QW18 : INT; q8 AT %QW20 : INT;
  END_VAR
  q0 := SHR(i, 1);
  q1 := SHR(i, 20);
  q2 := SHL(i, 2);
  q3 := ROL(INT#-32768, 1);
  q4 := SHR(u, n);
  b0 := d.0;
  b1 := d.1;
  d.0 := TRUE;
  q5 := d;
  k.%X15 := TRUE;
  q6 := k;
  q7 := REAL_TO_INT(EXPT(base, e));
  q8 := LREAL_TO_INT(EXPT(q, 3));
END_PROGRAM

CONFIGURATION cf
  RESOURCE r ON x
    TASK tk(INTERVAL := T#10ms, PRIORITY := 1);
    PROGRAM p WITH tk : main;
  END_RESOURCE
END_CONFIGURATION

(* ---- keptref.st ---- *)
(* A reference a RETAIN program instance keeps (W0006; Ed.3 6.5.6.2):
   kept as it is across a warm restart, as CODESYS and TwinCAT keep a
   pointer in retained memory; the plain instance's is NULL again.
   Worked by hand:

   tick 0: both take r := REF(x), n 1, and count through it: x 1 (Q0
   01 00, Q4 01 00; n Q2 01, Q6 01).
   tick 1: x 2, n stays 1.
   warm, before tick 2: a keeps r, x 2 and n 1; b starts again.
   tick 2: a counts on, x 3 (03 00), n 1; b takes the reference again,
   n 1, x 1.
   reference-skip: untried; the reference host has no warm restart. *)
PROGRAM main
  VAR r : REF_TO INT; x : INT; n : USINT; END_VAR
  VAR q AT %Q* : INT; qn AT %Q* : USINT; END_VAR
  IF r = NULL THEN
    r := REF(x);
    n := n + 1;
  END_IF;
  r^ := r^ + 1;
  q := x;
  qn := n;
END_PROGRAM
CONFIGURATION plant
  RESOURCE cpu ON PLC
    TASK t(INTERVAL := T#10ms, PRIORITY := 1);
    PROGRAM RETAIN a WITH t : main;
    PROGRAM b WITH t : main;
  END_RESOURCE
  VAR_CONFIG
    cpu.a.q AT %QW0 : INT;
    cpu.a.qn AT %QB2 : USINT;
    cpu.b.q AT %QW4 : INT;
    cpu.b.qn AT %QB6 : USINT;
  END_VAR
END_CONFIGURATION

(* ---- layout.st ---- *)
(* Structures with relative locations (Ed.3 6.4.4.7): each component at
   its byte, a BOOL at its bit, gaps between; OVERLAP lets components
   share bytes. The layout is iecf's (docs/c-output.md §4): little-endian,
   a structure the same bytes in C memory as at an address, an array or
   structure inside it back to back. Worked by hand:

   init: m (Com_data, %MB0..%MB25) has C1's initial values where C1 and
   C2 share bytes, C1 being declared first: length 26 at byte 2 (M 1a).
   q (Frame, %QB0..%QB15): id A5, pts 0, name 'ab' (61 62 00 00), byte 13
   lit (bit 7) 80, w BEEF (ef be).

   tick 0:
   c.C2.data2 := 1.0 puts 16#3F800000 at c's bytes 5 to 8 (00 00 80 3f);
   c.C1.head 16#1234 (34 12); c.C2.flag2 bit 3 and c.C1.flag1 bit 0 of
   byte 3 (09); length still 26. m := c: M 34 12 1a 09 00 00 00 80 3f,
   then 0. m.C2.data1 := 16#7F writes byte 5, data2's low byte (M5 7f);
   x := m.C2.data2 > 1.0 is TRUE, data2 16#3F80007F: %QX16.0.
   q.pts[1].y := -2: element 1 at byte 5, y 2 further, bytes 7, 8
   (fe ff); q.pts[0].act := TRUE, byte 2 (01). Bump(q.pts[1].y) adds 1
   through an in-out: -1 (ff ff). q.hi := q.lit: byte 13 81; Flip(q.hi)
   through an in-out: 80 again.
   f := q, the 16 bytes into C memory. f.id + 1: A6. f.name := 'xyz'
   (78 79 7a 00). ri := REF(f.pts[1].y); ri^ + 10: 9 (09 00).
   rb := REF(f.lit); rb^ := FALSE: byte 13 00. q := f: Q a6 00 01 00 00
   00 00 09 00 78 79 7a 00 00 ef be.
   r := REF(c1), a C pointer, r^.tail := 16#EE: c1's byte 25 through
   the structure's bytes. r := REF(m.C1), in the image: r^.length :=
   r^.length + 1: M2 1b. g := Make(16#11): a function's result, id 11,
   copied whole into %QB17..%QB32 with h := g.w = 16#BEEF (TRUE, %QX16.1)
   and k := c1.tail = 16#EE (TRUE, %QX16.2).
   %QB17.. g: 11 00 00 00 00 00 00 00 00 61 62 00 00 80 ef be.

   tick 1: q is as tick 0 left it. y -2, then -1, as before; but
   q.lit is FALSE now, so q.hi := q.lit is FALSE and Flip makes it
   TRUE: byte 13 01. f := q brings id A6, f.id + 1 is A7: Q a7 00 01 00
   00 00 00 09 00 78 79 7a 00 01 ef be. m is c's bytes again, length
   26, then + 1: 1b again.
   reference-skip: the reference compiler (Ed.2) has no relative
   locations. *)
TYPE
  Com1_data : STRUCT
    head   AT %B0   : INT;
    length AT %B2   : USINT := 26;
    flag1  AT %X3.0 : BOOL;
    tail   AT %B25  : BYTE;
  END_STRUCT;
  Com2_data : STRUCT OVERLAP
    head   AT %B0   : INT;
    length AT %B2   : USINT;
    flag2  AT %X3.3 : BOOL;
    data1  AT %B5   : BYTE;
    data2  AT %B5   : REAL;
    tail   AT %B19  : BYTE;
  END_STRUCT;
  Com_data : STRUCT OVERLAP
    C1 AT %B0 : Com1_data;
    C2 AT %B0 : Com2_data;
  END_STRUCT;
  Pt : STRUCT x : BYTE; act : BOOL; y : INT; END_STRUCT;
  Frame : STRUCT
    id   AT %B0    : USINT := 16#A5;
    pts  AT %B1    : ARRAY [0..1] OF Pt;
    name AT %B9    : STRING[3] := 'ab';
    lit  AT %X13.7 : BOOL := TRUE;
    hi   AT %X13.0 : BOOL;
    w    AT %W14   : WORD := 16#BEEF;
  END_STRUCT;
END_TYPE
FUNCTION Bump : INT
  VAR_IN_OUT v : INT; END_VAR
  v := v + 1;
  Bump := v;
END_FUNCTION
FUNCTION Flip : BOOL
  VAR_IN_OUT b : BOOL; END_VAR
  b := NOT b;
  Flip := b;
END_FUNCTION
FUNCTION Make : Frame
  VAR_INPUT k : USINT; END_VAR
  Make.id := k;
END_FUNCTION
PROGRAM main
  VAR
    c : Com_data;
    c1 : Com1_data;
    f : Frame;
    r : REF_TO Com1_data;
    rb : REF_TO BOOL;
    ri : REF_TO INT;
    n : INT;
    b : BOOL;
  END_VAR
  VAR
    m AT %MB0 : Com_data;
    q AT %QB0 : Frame;
    x AT %QX16.0 : BOOL;
    h AT %QX16.1 : BOOL;
    k AT %QX16.2 : BOOL;
    g AT %QB17 : Frame;
  END_VAR
  c.C2.data2 := 1.0;
  c.C1.head := 16#1234;
  c.C2.flag2 := TRUE;
  c.C1.flag1 := TRUE;
  m := c;
  m.C2.data1 := 16#7F;
  x := m.C2.data2 > 1.0;
  q.pts[1].y := -2;
  q.pts[0].act := TRUE;
  n := Bump(q.pts[1].y);
  q.hi := q.lit;
  b := Flip(q.hi);
  f := q;
  f.id := f.id + 1;
  f.name := 'xyz';
  ri := REF(f.pts[1].y);
  ri^ := ri^ + 10;
  rb := REF(f.lit);
  rb^ := FALSE;
  q := f;
  r := REF(c1);
  r^.tail := 16#EE;
  r := REF(m.C1);
  r^.length := r^.length + 1;
  g := Make(16#11);
  h := g.w = 16#BEEF;
  k := c1.tail = 16#EE;
END_PROGRAM
CONFIGURATION plant
  RESOURCE r ON PLC
    TASK t (INTERVAL := T#10ms, PRIORITY := 1);
    PROGRAM p WITH t : main;
  END_RESOURCE
END_CONFIGURATION

(* ---- ldates.st ---- *)
(* LDATE, LTOD and LDT (Ed.3 Table 10, 22, 30, 36; docs/dependencies.md):
   signed 64-bit nanoseconds, LDT from 1677-09-21 to 2262-04-11. An LTOD
   and an LDT go on 7 hours a tick, from LTOD#20:00:00.000000001 and
   LDT#1969-12-31-20:00:00.5; each tick shows, as bits, comparisons of
   what the operators, conversions and Table 36 give. An LTOD wraps at
   midnight; a long value made a short one rounds down. iecf only
   (reference-skip: the reference compiler has no L dates). *)
PROGRAM main
VAR
  r_bits AT %MW0 : WORD;
  r_year AT %MW2 : UINT;
  r_ms AT %MW4 : UINT;
END_VAR
VAR
  clock : LTOD := LTOD#20:00:00.000_000_001;
  stamp : LDT := LDT#1969-12-31-20:00:00.5;
  start : LDT := LDT#1969-12-31-00:00:00;
  day : LDATE;
  span : LTIME;
  mo, da, h, mi, s : UINT;
END_VAR
clock := clock + T#7h;
stamp := ADD_LDT_LTIME(stamp, LTIME#7h);
day := LDT_TO_LDATE(stamp);
span := T#1500ms;
r_bits := 0;
IF clock < LTOD#12:00:00 THEN r_bits := r_bits OR 16#0001; END_IF;
IF LDT_TO_LTOD(stamp) - clock = LTIME#499_999_999ns THEN r_bits := r_bits OR 16#0002; END_IF;
IF stamp - start > LTIME#1d THEN r_bits := r_bits OR 16#0004; END_IF;
IF SUB_LTOD_LTOD(LTOD#01:00:00, LTOD#23:00:00) = LTIME#-22h THEN r_bits := r_bits OR 16#0008; END_IF;
IF CONCAT_DATE_LTOD(LDT_TO_DATE(stamp), LDT_TO_LTOD(stamp)) = stamp THEN r_bits := r_bits OR 16#0010; END_IF;
IF LDT_TO_LDATE(LDT#1969-12-31-23:59:59.999999999) = LD#1969-12-31 THEN r_bits := r_bits OR 16#0020; END_IF;
IF LDT_TO_DT(stamp) = DT#1970-01-01-03:00:00 THEN r_bits := r_bits OR 16#0040; END_IF;
IF SUB_LDT_LTIME(stamp, LTIME#1d) < start THEN r_bits := r_bits OR 16#0080; END_IF;
IF LTOD_TO_TOD(clock) = TOD#03:00:00 THEN r_bits := r_bits OR 16#0100; END_IF;
IF LTIME_TO_TIME(LTIME#-1500us) = T#-2ms THEN r_bits := r_bits OR 16#0200; END_IF;
IF span = LTIME#1500ms THEN r_bits := r_bits OR 16#0400; END_IF;
IF DT_TO_LDT(DT#2026-11-08-12:00:00) = LDT#2026-11-08-12:00:00 THEN r_bits := r_bits OR 16#0800; END_IF;
IF clock - LTIME#21h = LTOD#06:00:00.000000001 THEN r_bits := r_bits OR 16#1000; END_IF;
IF STRING_TO_LDT(LDT_TO_STRING(stamp)) = stamp THEN r_bits := r_bits OR 16#2000; END_IF;
IF MAX(stamp, start) = stamp THEN r_bits := r_bits OR 16#4000; END_IF;
IF day = LD#1970-01-02 THEN r_bits := r_bits OR 16#8000; END_IF;
SPLIT_LDT(LDT#1677-09-21-00:12:43.145224192, r_year, mo, da, h, mi, s, r_ms);
END_PROGRAM

CONFIGURATION plant
  RESOURCE r ON PLC
    TASK fast(INTERVAL := T#10ms, PRIORITY := 0);
    PROGRAM p WITH fast : main;
  END_RESOURCE
END_CONFIGURATION

(* ---- leftout.st ---- *)
(* A standard function called by name with inputs left out (Ed.3
   6.6.1.4.2: "Any variable to which no value is assigned in the list
   shall have ... the default value for the associated data type"):
   each takes its type's default, 0, FALSE, '' or D#1970-01-01. An
   extensible function has as many inputs as the highest name given
   (6.6.2.5.1); those below it not given are left out. Worked by hand,
   the same at every tick, v 7, m -2, t TRUE, w 16#00F0:
   LIMIT(IN := v, MX := 5) 5, MN 0 (Table 19, NOTE 3) (%QB0);
   LIMIT(IN := m, MX := 5) 0 (%QB1); MUL(IN2 := v) 0 * 7 = 0 (%QB2);
   MAX(IN2 := m) 0 (%QB3); MIN(IN2 := v) 0 (%QB4); SUB(IN2 := v) -7
   (%QB5); MUX_INT(K := 3, IN0 := 1, IN2 := 2, IN4 := 3) 0, IN3 left out
   (6.6.2.5.1, EXAMPLE 2) (%QB6); SEL(G := t, IN0 := v) 0 (%QB7);
   ADD(IN3 := v) 0 + 0 + 7 = 7 (%QB8); the constant k, LIMIT(IN := 9,
   MX := 5), 5 (%QB9). AND(IN2 := t) FALSE (%QX10.0); OR(IN3 := t) TRUE
   (%QX10.1); XOR(IN2 := t) TRUE (%QX10.2); GT(IN3 := m) 0 > 0 > -2
   FALSE (%QX10.3); GT(IN2 := m) 0 > -2 TRUE (%QX10.4); EQ(IN2 := 0) TRUE
   (%QX10.5); SHL(IN := w) w (%QX10.6); LEN() 0 (%QX10.7).
   LEFT(IN := 'abc') '' (%QX11.0); DELETE(IN := 'abc', P := 2) 'abc',
   L 0 (%QX11.1); INSERT(IN1 := 'ab', P := 1) 'ab' (%QX11.2);
   CONCAT(IN2 := 'x') 'x' (%QX11.3); FIND(IN1 := 'abc') 0 (%QX11.4);
   EXPT(IN1 := 2.0) 1.0 (%QX11.5); CONCAT_TOD(HOUR := 1) TOD#01:00:00
   (%QX11.6); DINT_TO_INT() 0 (%QX11.7). SPLIT_DATE(YEAR => y) of
   D#1970-01-01: y 1970 (%QW12, 16#07B2).
   reference-skip: the reference compiler's C for an extensible function
   called by name without IN1, MUL(IN2 := v), does not compile (too few
   arguments); it has no LEN() or DINT_TO_INT() without an input, no
   MUX_INT, none of Table 36's. *)
PROGRAM main
  VAR
    v : INT := 7;
    m : INT := -2;
    t : BOOL := TRUE;
    w : WORD := 16#00F0;
    s : STRING;
    r : REAL;
    td : TOD;
    y : UINT;
  END_VAR
  VAR CONSTANT
    k : INT := LIMIT(IN := 9, MX := 5);
  END_VAR
  VAR
    q0 AT %QB0 : SINT;
    q1 AT %QB1 : SINT;
    q2 AT %QB2 : SINT;
    q3 AT %QB3 : SINT;
    q4 AT %QB4 : SINT;
    q5 AT %QB5 : SINT;
    q6 AT %QB6 : SINT;
    q7 AT %QB7 : SINT;
    q8 AT %QB8 : SINT;
    q9 AT %QB9 : SINT;
    b0 AT %QX10.0 : BOOL;
    b1 AT %QX10.1 : BOOL;
    b2 AT %QX10.2 : BOOL;
    b3 AT %QX10.3 : BOOL;
    b4 AT %QX10.4 : BOOL;
    b5 AT %QX10.5 : BOOL;
    b6 AT %QX10.6 : BOOL;
    b7 AT %QX10.7 : BOOL;
    c0 AT %QX11.0 : BOOL;
    c1 AT %QX11.1 : BOOL;
    c2 AT %QX11.2 : BOOL;
    c3 AT %QX11.3 : BOOL;
    c4 AT %QX11.4 : BOOL;
    c5 AT %QX11.5 : BOOL;
    c6 AT %QX11.6 : BOOL;
    c7 AT %QX11.7 : BOOL;
    qy AT %QW12 : UINT;
  END_VAR
  q0 := INT_TO_SINT(LIMIT(IN := v, MX := 5));
  q1 := INT_TO_SINT(LIMIT(IN := m, MX := 5));
  q2 := INT_TO_SINT(MUL(IN2 := v));
  q3 := INT_TO_SINT(MAX(IN2 := m));
  q4 := INT_TO_SINT(MIN(IN2 := v));
  q5 := INT_TO_SINT(SUB(IN2 := v));
  q6 := INT_TO_SINT(MUX_INT(K := v - 4, IN0 := 1, IN2 := 2, IN4 := 3));
  q7 := INT_TO_SINT(SEL(G := t, IN0 := v));
  q8 := INT_TO_SINT(ADD(IN3 := v));
  q9 := INT_TO_SINT(k);
  b0 := AND(IN2 := t);
  b1 := OR(IN3 := t);
  b2 := XOR(IN2 := t);
  b3 := GT(IN3 := m);
  b4 := GT(IN2 := m);
  b5 := EQ(IN2 := 0);
  b6 := SHL(IN := w) = w;
  b7 := LEN() = 0;
  s := 'abc';
  c0 := LEFT(IN := s) = '';
  c1 := DELETE(IN := s, P := 2) = 'abc';
  c2 := INSERT(IN1 := 'ab', P := 1) = 'ab';
  c3 := CONCAT(IN2 := 'x') = 'x';
  c4 := FIND(IN1 := s) = 0;
  r := 2.0;
  c5 := EXPT(IN1 := r) = 1.0;
  td := CONCAT_TOD(HOUR := 1);
  c6 := td = TOD#01:00:00;
  c7 := DINT_TO_INT() = 0;
  SPLIT_DATE(YEAR => y);
  qy := y;
END_PROGRAM

CONFIGURATION c
  RESOURCE r ON x
    TASK t(INTERVAL := T#10ms, PRIORITY := 1);
    PROGRAM p WITH t : main;
  END_RESOURCE
END_CONFIGURATION

(* ---- litcalls.st ---- *)
(* A standard function given literals alone, and a quotient of real
   literals: no operand gives the expression a type, so it is computed
   in the type wanted of it - the variable assigned, the other operand,
   the conversion's own. Worked by hand, the same at every tick:
   v := MAX(10, 11): 11 (%QB0). r := SQRT(2.0), 1.4142135, times 10.0:
   14 (%QB1). SEL(TRUE, 1, 2): 2 (%QB2). w := SHL(1, 3): 8 (%QB3).
   ABS(-3): 3 (%QB4). r := 1.0 / 3.0, times 9.0: 3 (%QB5).
   LIMIT(1, 5, 3): 3 (%QB6). MUX(1, 5, 6), the second of its inputs: 6
   (%QB7). ADD(1, 2, 3): 6 (%QB8). r := MAX(1.5, 2), times 2.0: 4
   (%QB9). v := 10; v := v + MAX(1, 2): 12 (%QB10).
   Integers stay integers where a real is wanted: r := MAX(7, 2) / 2 is
   7 / 2, 3, as r := 7 / 2 is (%QB16): times 2.0, 6 (%QB11); r := 1.5 +
   7 / 2 is 4.5: times 2.0, 9 (%QB12).
   -MAX(1, 2): -2 (%QB13). GT(MAX(1, 2), 1): TRUE (%QX14.0).
   REAL_TO_INT(SQRT(16.0)): 4 (%QB15). d := ADD(30000, 30000) in DINT:
   60000, over 1000 is 60 (%QB17). lr := SQRT(2.0) in LREAL: lr * lr *
   50.0 is 100.00000000000001, 100 (%QB18). COS(0): 1 (%QB19).
   EXPT(2.0, 3): 8 (%QB20). (MAX(1, 2)) + 1: 3 (%QB21).
   An initial value: i : INT := MAX(1, 2), 2 (%QB23).
   Last, the same ADD(30000, 30000) wanted as an INT is computed in
   INT: it wraps to -5536 and is flagged OVERFLOW; over 100 is -55
   (%QB22).
   reference-skip: a function call in an initial value: the reference
   compiler refuses it. *)
PROGRAM main
  VAR
    v : INT;
    r : REAL;
    lr : LREAL;
    b : BOOL;
    w : WORD;
    d : DINT;
    i : INT := MAX(1, 2);
  END_VAR
  VAR
    q0 AT %QB0 : SINT;
    q1 AT %QB1 : SINT;
    q2 AT %QB2 : SINT;
    q3 AT %QB3 : SINT;
    q4 AT %QB4 : SINT;
    q5 AT %QB5 : SINT;
    q6 AT %QB6 : SINT;
    q7 AT %QB7 : SINT;
    q8 AT %QB8 : SINT;
    q9 AT %QB9 : SINT;
    q10 AT %QB10 : SINT;
    q11 AT %QB11 : SINT;
    q12 AT %QB12 : SINT;
    q13 AT %QB13 : SINT;
    q14 AT %QX14.0 : BOOL;
    q15 AT %QB15 : SINT;
    q16 AT %QB16 : SINT;
    q17 AT %QB17 : SINT;
    q18 AT %QB18 : SINT;
    q19 AT %QB19 : SINT;
    q20 AT %QB20 : SINT;
    q21 AT %QB21 : SINT;
    q22 AT %QB22 : SINT;
    q23 AT %QB23 : SINT;
  END_VAR
  v := MAX(10, 11);
  q0 := INT_TO_SINT(v);
  r := SQRT(2.0);
  q1 := REAL_TO_SINT(r * 10.0);
  v := SEL(TRUE, 1, 2);
  q2 := INT_TO_SINT(v);
  w := SHL(1, 3);
  q3 := WORD_TO_SINT(w);
  v := ABS(-3);
  q4 := INT_TO_SINT(v);
  r := 1.0 / 3.0;
  q5 := REAL_TO_SINT(r * 9.0);
  v := LIMIT(1, 5, 3);
  q6 := INT_TO_SINT(v);
  v := MUX(1, 5, 6);
  q7 := INT_TO_SINT(v);
  v := ADD(1, 2, 3);
  q8 := INT_TO_SINT(v);
  r := MAX(1.5, 2);
  q9 := REAL_TO_SINT(r * 2.0);
  v := 10;
  v := v + MAX(1, 2);
  q10 := INT_TO_SINT(v);
  r := MAX(7, 2) / 2;
  q11 := REAL_TO_SINT(r * 2.0);
  r := 1.5 + 7 / 2;
  q12 := REAL_TO_SINT(r * 2.0);
  v := -MAX(1, 2);
  q13 := INT_TO_SINT(v);
  q14 := GT(MAX(1, 2), 1);
  v := REAL_TO_INT(SQRT(16.0));
  q15 := INT_TO_SINT(v);
  r := 7 / 2;
  q16 := REAL_TO_SINT(r);
  d := ADD(30000, 30000);
  q17 := DINT_TO_SINT(d / 1000);
  lr := SQRT(2.0);
  q18 := LREAL_TO_SINT(lr * lr * 50.0);
  r := COS(0);
  q19 := REAL_TO_SINT(r);
  r := EXPT(2.0, 3);
  q20 := REAL_TO_SINT(r);
  v := (MAX(1, 2)) + 1;
  q21 := INT_TO_SINT(v);
  q23 := INT_TO_SINT(i);
  v := ADD(30000, 30000);
  q22 := INT_TO_SINT(v / 100);
END_PROGRAM

CONFIGURATION c
  RESOURCE r ON x
    TASK t(INTERVAL := T#10ms, PRIORITY := 1);
    PROGRAM p WITH t : main;
  END_RESOURCE
END_CONFIGURATION

(* ---- located.st ---- *)
(* Variables at an address (Ed.3 6.5.5.3; docs/c-output.md §4): the
   address is where a variable starts, and it takes its own type's width
   from there, little-endian - a TIME, DATE or TOD 4 bytes, an LTIME or
   LDT 8, whatever the size prefix says (W0004 when it differs). A BOOL
   at a byte takes the whole byte: TRUE written as 1, any value but 0
   read as TRUE. A program's TIME output connected to an LTIME global at
   an address is converted, ms to ns. iecf only (reference-skip: the
   reference compiler refuses an LTIME at an address, and holds a TIME,
   DATE, TOD or DT as a structure of seconds and nanoseconds, not 4
   bytes). *)
PROGRAM main
VAR_INPUT
  tick : TIME;
END_VAR
VAR_OUTPUT
  el_out : TIME;
END_VAR
VAR
  el AT %MD0 : TIME;
  big AT %ML4 : LTIME;
  day AT %MD12 : DATE;
  odd AT %MW16 : TIME;
  r AT %MB20 : REAL;
  toggle AT %QB0 : BOOL;
  seen AT %QX1.0 : BOOL;
  inb AT %IB0 : BOOL;
END_VAR
VAR
  n : INT;
END_VAR
n := n + 1;
el := el - tick;
big := el;
IF n = 2 THEN day := D#2026-11-08; END_IF;
odd := el + T#1ms;
r := INT_TO_REAL(n) / 2.0;
toggle := NOT toggle;
seen := inb;
el_out := el;
END_PROGRAM

CONFIGURATION plant
  VAR_GLOBAL
    g AT %ML24 : LTIME;
  END_VAR
  RESOURCE r ON PLC
    TASK fast(INTERVAL := T#10ms, PRIORITY := 0);
    PROGRAM p WITH fast : main(tick := T#250ms, el_out => g);
  END_RESOURCE
END_CONFIGURATION

(* ---- locinit.st ---- *)
(* The initial value of a variable at an address that its type gives
   without the declaration saying so (Ed.3 6.4.4.2.2, 6.4.4.4.2): an
   enumeration starts at its first value, a subrange at its lower limit,
   and a structure or array holding them likewise. Until 2026-11-13 these
   were left at 0 when no initial value was written out. Worked by hand:

   init: e (Mode, first value Run = 5) at %QW0: 05 00; lim, SINT(3..5),
   at %QB2: 03; h, a Hold (m Mode, s SINT(-2..2)), at %QW3: 05 00 fe;
   arr, two Mode at %QW6: 05 00 05 00; zero, SINT(0..9) at %QB10 starts
   at 0: 00. ein, a Mode at %IW0, is the platform's: not written, and
   so ein = Run is FALSE: %QB11 00 at tick 0.
   tick 0: e := Halt (06 00); the rest as at init.
   reference-skip: enumerated values, arrays and structures at an
   address: refused. *)
TYPE
  Mode : (Run := 5, Halt);
  Hold : STRUCT m : Mode; s : SINT(-2..2); END_STRUCT;
END_TYPE
PROGRAM main
  VAR
    e AT %QW0 : Mode;
    lim AT %QB2 : SINT(3..5);
    h AT %QW3 : Hold;
    arr AT %QW6 : ARRAY [0..1] OF Mode;
    zero AT %QB10 : SINT(0..9);
    copy AT %QB11 : BYTE;
  END_VAR
  VAR
    ein AT %IW0 : Mode;
  END_VAR
  copy := BOOL_TO_BYTE(ein = Run);
  e := Halt;
END_PROGRAM
CONFIGURATION plant
  RESOURCE r ON PLC
    TASK t (INTERVAL := T#10ms, PRIORITY := 1);
    PROGRAM p WITH t : main;
  END_RESOURCE
END_CONFIGURATION

(* ---- loopflag.st ---- *)
(* One statement's overflow carried across a FOR loop (runtime/iecf.h
   iecf_*_or, crates/iecf-codegen stmt.rs loop_flags): the loop's only
   statement that can flag ORs its overflow into a local, taken after the
   loop with its line; the FOR's own step is taken after that. The order
   is the run's. Worked by hand:
   tick 0: x 2147483000, plus 100 on each of i = 32760..32767, eight
   passes: the seventh leaves DINT (2147483700): wrapped, flagged at
   x := x + 100 (line 23), the first flag. x ends 2147483800 - 2^32 =
   -2147483496 (MD2 98 00 00 80). The FOR's step past 32767 leaves INT
   too, flagged after (not the first): i -32768 (MW0 00 80), n := i
   (MW6 00 80).
   tick 1: the same; the first flag stays.
   reference-skip: the reference compiler's FOR to INT's last value does
   not end (its counter wraps). *)
PROGRAM main
VAR
  i AT %MW0 : INT;
  x AT %MD2 : DINT;
  n AT %MW6 : INT;
END_VAR
x := 2147483000;
FOR i := 32760 TO 32767 DO
  x := x + 100;
END_FOR;
n := i;
END_PROGRAM

CONFIGURATION Plant
  RESOURCE R ON PLC
    TASK fast(INTERVAL := T#10ms, PRIORITY := 1);
    PROGRAM P WITH fast : main;
  END_RESOURCE
END_CONFIGURATION

(* ---- loopflag2.st ---- *)
(* As loopflag, the statement never overflowing: x 0, plus 100 on each of
   eight passes, 800 (MD2 20 03 00 00). The FOR's step past 32767 is the
   only flag, at the FOR's line (13): i -32768 (MW0 00 80), n -32768.
   reference-skip: the reference compiler's FOR to INT's last value does
   not end (its counter wraps). *)
PROGRAM main
VAR
  i AT %MW0 : INT;
  x AT %MD2 : DINT;
  n AT %MW6 : INT;
END_VAR
x := 0;
FOR i := 32760 TO 32767 DO
  x := x + 100;
END_FOR;
n := i;
END_PROGRAM

CONFIGURATION Plant
  RESOURCE R ON PLC
    TASK fast(INTERVAL := T#10ms, PRIORITY := 1);
    PROGRAM P WITH fast : main;
  END_RESOURCE
END_CONFIGURATION

(* ---- narrow.st ---- *)
(* A narrowing conversion out of the target's range keeps the low bits,
   as CODESYS and TwinCAT have it (INT_TO_SINT(4223) = 127), and the reference compiler's
   C cast does; iecf also flags it (PROPOSAL.md §6.3). At tick 1, 4223
   leaves SINT: both give 127, and iecf records "flag 4 MAIN 18" in
   ctx->flag. At tick 2, -1 leaves UINT: 65535. Its trace is
   narrow.iecf.trace: the reference compiler's bytes, with the flag from tick 1. *)
PROGRAM main
VAR
  a AT %IW0 : INT;
  s AT %MB0 : SINT;
  u AT %MW2 : UINT;
END_VAR
VAR
  d : DINT;
END_VAR
d := INT_TO_DINT(a);
u := DINT_TO_UINT(d);
s := INT_TO_SINT(a);
END_PROGRAM

CONFIGURATION plant
  RESOURCE r ON PLC
    TASK fast(INTERVAL := T#10ms, PRIORITY := 0);
    PROGRAM p WITH fast : main;
  END_RESOURCE
END_CONFIGURATION

(* ---- narrowing.st ---- *)
(* implicit-narrowing: an integer or bit string where another is wanted,
   converted as its *_TO_* would, W0010 at each. Worked by hand:
   i := d, DINT 100000 (16#186A0) into an INT: its low 16 bits, 16#86A0,
   -31072, flagged (%QW0).
   w := m, INT -2 into a WORD: its bits, 16#FFFE, unflagged (%QW2).
   u := m, INT -2 into a UINT: low bits, 65534, flagged (%QW4).
   g(i), the INT -31072 passed to a SINT input: low 8 bits 16#A0, -96,
   flagged (%QB6).
   q4 := b, BYTE 200 into an INT: 200, which it holds (%QW8).
   The first flag is i := d's, line 28.
   reference-skip: implicit narrowing is CODESYS's, not IEC 61131-3. *)
FUNCTION g : SINT
  VAR_INPUT x : SINT; END_VAR
  g := x;
END_FUNCTION

PROGRAM main
  VAR
    i : INT; d : DINT := 100000; w : WORD; u : UINT; m : INT := -2; b : BYTE := 200;
  END_VAR
  VAR
    q0 AT %QW0 : INT;
    q1 AT %QW2 : WORD;
    q2 AT %QW4 : UINT;
    q3 AT %QB6 : SINT;
    q4 AT %QW8 : INT;
  END_VAR
  i := d;
  q0 := i;
  w := m;
  q1 := w;
  u := m;
  q2 := u;
  q3 := g(i);
  q4 := b;
END_PROGRAM

CONFIGURATION cf
  RESOURCE r ON x
    TASK tk(INTERVAL := T#10ms, PRIORITY := 1);
    PROGRAM p WITH tk : main;
  END_RESOURCE
END_CONFIGURATION
